(* IEC 61131-3 sources: daoli-st-library/DL_Algo (part 8) *)

(* ---- FB_DL_AutoTuneRelay.st ---- *)
(*
    FB_DL_AutoTuneRelay —— 继电反馈自整定
    ------------------------------------------------------------------
    分类      : DL_Algo / ControlLaw
    前缀      : FB_DL_
    版本      : 1.0.0
    溯源      : 公开学术判据 —— 继电反馈法（Astrom & Hagglund 1984）描述函数
                N(a) = 4d/(pi*a)，含迟滞时 -1/N(a) = -(pi/4d)*sqrt(a^2 - h^2)；
                整定规则取 Ziegler-Nichols 与 Astrom-Hagglund 公开文本；
                只借公开公式与规则常数（属公共知识），测量闸门、状态机、引脚契约与
                码位 100% 自有；clean-room 重写，未复制任何闭源厂商源码
    平台      : 纯 IEC 61131-3，CODESYS V3.5+ / TwinCAT 3 / InoProShop 通用
    作者      : 道莅代码库 · PLC编程专家（R19）
    ------------------------------------------------------------------
    功能说明  : 把 ±d 继电（可带迟滞 h）接入回路，等振幅稳定后测极限振荡周期 Tu 与幅值 a，
                按公开描述函数算临界增益 Ku，再按选定规则给出 Kp / Ti / Td。
                本件不闭环控制，只输出 bRelayOut（接上层手动通道）与整定结果。
                核心防御：① 继电幅值非正/非有限即故障级 2A10（d = 0 时 Ku = 0，结果无意义）；
                ② 迟滞不小于实测幅值时拒绝出结果（描述函数分母为零/虚数，Ku 不可定义）；
                ③ 每半周期采样数不足即故障级 2A11——采样太疏时测出的「振荡」是采样网格
                   产物，不是对象特性（R67 采样密度闸先行）；
                ④ 幅值稳定判据不通过只置信息码继续测，超时才是故障级 2A12；
                ⑤ bAbort 必须撤继电（本件最高危点：不撤则回路一直振荡），且人为中止不置故障。
                说明：继电幅值相对满量程 20% 的工程上限需满量程信息，本件无满量程引脚，
                该上限由调用方在上层保证（头注释留档，不做无法判定的检查）。
    错误码    : 16#0002_2A01 振荡未收敛，继续测量 / 参数超域已钳位——信息级，正常防御
                16#0002_2A02 预留禁用（信息级，不得挪用）
                16#0002_2A10 继电参数非法（d 非正或非有限、h >= a、采样周期越域）——故障级，中止实验并撤继电
                16#0002_2A11 半周期采样密度不足，振荡不可信——故障级，中止实验并撤继电
                16#0002_2A12 超时未收敛 / Ku 不可表示 / 整定规则落 ELSE 兜底——故障级，中止实验并撤继电
    码位总账  : 16#0002_2A01 用 / 16#0002_2A02 预留 ｜ 16#0002_2A10 用 / 16#0002_2A11 用 / 16#0002_2A12 用
    状态机    : E_DL_TuneState（eIdle / eRelay / eMeasure / eDone / eFault）五态，CASE 含 ELSE 兜底，
                ELSE 回 eIdle 并置故障级 2A12；bAbort 沿无条件回 eIdle 且撤继电。
    采样约定  : fbTrigStart / fbTrigAbort / fbTimeout 在本体首部无条件刷新，绝不放入 IF 或 CASE；
                时间基准由 tSampleTime 引脚累加，累加前用比较式预判溢出（不靠回绕兜底）；
                整定规则按公开文本：ZN-P 0.5Ku；ZN-PI 0.45Ku / Tu*1.2^-1；ZN-PID 0.6Ku / Tu/2 / Tu/8；
                AH 无超调 0.2Ku / Tu/2 / Tu/3。
    修订记录  : 2026-11-16 v1.0.0 首次入库（R19）
*)

(*
    枚举 : E_DL_TuneRule —— 整定规则（本文件为全库唯一属主）
*)
TYPE E_DL_TuneRule :
(
    eZnP           := 0,                      // Ziegler-Nichols 纯比例规则 / Ziegler-Nichols proportional rule
    eZnPi          := 1,                      // Ziegler-Nichols 比例积分规则 / Ziegler-Nichols PI rule
    eZnPid         := 2,                      // Ziegler-Nichols 比例积分微分规则 / Ziegler-Nichols PID rule
    eAhNoOvershoot := 3                       // Astrom-Hagglund 无超调规则 / Astrom-Hagglund no overshoot rule
);
END_TYPE

(*
    枚举 : E_DL_TuneState —— 自整定实验状态（本文件为全库唯一属主）
*)
TYPE E_DL_TuneState :
(
    eIdle    := 0,                            // 空闲：继电输出撤销 / idle, relay output withdrawn
    eRelay   := 1,                            // 施加继电，等待首个翻转 / relay applied, waiting for the first flip
    eMeasure := 2,                            // 收集中：测幅值与半周期 / measuring amplitude and half periods
    eDone    := 3,                            // 完成：结果有效 / done, results valid
    eFault   := 4                             // 故障：实验中止 / fault, experiment aborted
);
END_TYPE

FUNCTION_BLOCK FB_DL_AutoTuneRelay
VAR_INPUT
    bEnable           : BOOL;                 // 使能，FALSE 中止实验并撤继电 / enable, FALSE aborts the experiment and withdraws the relay
    bStart            : BOOL;                 // 启动，上升沿启动实验（运行中忽略）/ start, rising edge begins the experiment, ignored while running
    bAbort            : BOOL;                 // 中止，上升沿中止并回 eIdle（不置故障）/ abort, rising edge aborts back to idle without raising a fault
    fPv               : REAL := 0.0;          // 过程测量（被控量）[用户单位] / process measurement [user unit]
    fSp               : REAL := 0.0;          // 目标值，实验围绕此点进行 [用户单位] / setpoint the experiment oscillates around [user unit]
    fRelayAmp         : REAL := 5.0;          // 继电幅值 d [用户单位]，必须 > 0 / relay amplitude d [user unit], must be > 0
    fRelayHyst        : REAL := 0.2;          // 继电迟滞 h [用户单位]，范围 0.0~fRelayAmp（含等号即非法）/ relay hysteresis h [user unit], 0.0~fRelayAmp, equality is illegal
    uCyclesRequired   : UINT := 4;            // 需要观察的完整振荡周期数 [周期]，范围 2~20 / number of full cycles to observe [cycle], range 2~20
    uMinSamplesPerHalf : UINT := 6;           // 每半周期最少采样数 [拍]，范围 4~100 / minimum samples per half period [scan], range 4~100
    tMaxDuration      : TIME := T#300S;       // 实验总超时 [ms]，范围 10 s~2 h / experiment timeout [ms], range 10 s~2 h
    fStabTolPercent   : REAL := 2.0;          // 幅值稳定判据：前后半窗均值差百分比上限 [%]，范围 0.1~20.0 / amplitude stability tolerance [%], range 0.1~20.0
    eRule             : E_DL_TuneRule := eZnPid; // 整定规则 / tuning rule
    tSampleTime       : TIME := T#100MS;      // 采样周期 [ms]，范围 1~10000 / sample time [ms], range 1~10000
END_VAR
VAR_OUTPUT
    bRelayOut         : BOOL;                 // 继电输出（TRUE = 加 +d），接上层手动通道 / relay output, TRUE adds plus d, wired to the manual channel
    bBusy             : BOOL;                 // 实验进行中 / experiment running
    bDone             : BOOL;                 // 完成（单周期脉冲，结果有效）/ done, single-cycle pulse with valid results
    fOscAmp           : REAL;                 // 测得振荡幅值 a [用户单位] / measured oscillation amplitude a [user unit]
    tUltPeriod        : TIME;                 // 测得极限周期 Tu [ms] / measured ultimate period Tu [ms]
    fUltGain          : REAL;                 // 临界增益 Ku [无量纲] / ultimate gain Ku [dimensionless]
    fKp               : REAL;                 // 整定比例增益 [无量纲] / tuned proportional gain [dimensionless]
    fTi               : REAL;                 // 整定积分时间 [s]，0 表示纯 P / tuned integral time [s], zero means pure P
    fTd               : REAL;                 // 整定微分时间 [s]，0 表示无微分 / tuned derivative time [s], zero means no derivative
    uCycleDone        : UINT;                 // 已完成的有效振荡周期数 [周期] / completed valid cycles [cycle]
    eErr              : UDINT;                // 错误码，0=正常 / error id, 0=ok
    bError            : BOOL;                 // 故障标志，eErr 为故障级时 TRUE / error flag, TRUE on fault-level eErr
    bValid            : BOOL;                 // 结果是否可用 / results valid flag
END_VAR
VAR
    eState            : E_DL_TuneState := eIdle; // 状态机当前态 / current state machine state
    fbTrigStart       : R_TRIG;               // 启动沿实例，本体首部无条件刷新 / start edge instance, refreshed unconditionally
    fbTrigAbort       : R_TRIG;               // 中止沿实例，本体首部无条件刷新 / abort edge instance, refreshed unconditionally
    fbTimeout         : TON;                  // 实验总超时实例，本体首部无条件刷新 / total timeout instance, refreshed unconditionally
    bRelayPrev        : BOOL;                 // 上一拍继电输出，翻转检测用 / previous relay output for flip detection
    fPeakHi           : REAL;                 // 本半周期上峰值 [用户单位] / upper peak of the current half period [user unit]
    fPeakLo           : REAL;                 // 本半周期下峰值 [用户单位] / lower peak of the current half period [user unit]
    tNow              : TIME;                 // 实验内累计时间 [ms] / accumulated experiment time [ms]
    tEdgeLast         : TIME;                 // 上一次翻转的时刻 [ms] / time of the previous flip [ms]
    tHalf             : TIME;                 // 最近一个半周期长度 [ms] / most recent half period length [ms]
    tHalfPrev         : TIME;                 // 上一个半周期长度 [ms] / previous half period length [ms]
    uHalfCount        : UINT;                 // 已采集的半周期数 [个] / collected half periods [count]
    fAmpSum1          : REAL;                 // 第一窗幅值累计 [用户单位] / first window amplitude sum [user unit]
    fAmpSum2          : REAL;                 // 第二窗幅值累计 [用户单位] / second window amplitude sum [user unit]
    uAmpCnt1          : UINT;                 // 第一窗样本数 [个] / first window sample count [count]
    uAmpCnt2          : UINT;                 // 第二窗样本数 [个] / second window sample count [count]
    fHalfAmp          : REAL;                 // 单个半周期的幅值 [用户单位] / amplitude of one half period [user unit]
    fMean1            : REAL;                 // 第一窗均值 [用户单位] / first window mean [user unit]
    fMean2            : REAL;                 // 第二窗均值 [用户单位] / second window mean [user unit]
    fRelAmp           : REAL;                 // 幅值相对偏差 [无量纲] / relative amplitude deviation [dimensionless]
    fStabTolEff       : REAL;                 // 钳位后的稳定容差 [%] / clamped stability tolerance [%]
    fCyclesEff        : REAL;                 // 钳位后的周期数（REAL 形态，除法用）/ clamped cycle count in REAL form, used for division
    fHystEff          : REAL;                 // 钳位后的继电迟滞 [用户单位] / clamped relay hysteresis [user unit]
    fKuL              : LREAL;                // 临界增益中间量（LREAL 承载）/ ultimate gain intermediate carried in LREAL
    fAmpL             : LREAL;                // 幅值中间量（LREAL 承载）/ amplitude intermediate carried in LREAL
    fHystL            : LREAL;                // 迟滞中间量（LREAL 承载）/ hysteresis intermediate carried in LREAL
    fDenL             : LREAL;                // 描述函数分母（LREAL 承载）/ describing function denominator in LREAL
    fTuSec            : REAL;                 // 极限周期的秒值 [s] / ultimate period in seconds [s]
    nSampHalf         : DINT;                 // 单半周期采样数 [拍] / samples in one half period [scan]
    nDtMs             : DINT;                 // 采样周期毫秒整数 [ms] / sample time in integer milliseconds [ms]
    uNeedHalf         : UINT;                 // 需要采集的半周期总数 [个] / required half periods [count]
    bNonFin           : BOOL;                 // 输入非有限判定标志 / non-finite input flag
    bCollect          : BOOL;                 // 本拍完成一次有效半周期采集 / a valid half period was collected in this cycle
    uMinSampEff       : UINT;                 // 钳位后的每半周期最少采样数 [拍] / clamped minimum samples per half [scan]
END_VAR
VAR CONSTANT
    DL_AT_MIN_CYCLES    : UINT := 2;          // 周期数下限 [周期] / cycle count lower bound [cycle]
    DL_AT_MAX_CYCLES    : UINT := 20;         // 周期数上限 [周期] / cycle count upper bound [cycle]
    DL_AT_MIN_SAMPLES   : UINT := 4;          // 每半周期采样数下限 [拍] / samples per half lower bound [scan]
    DL_AT_MAX_SAMPLES   : UINT := 100;        // 每半周期采样数上限 [拍] / samples per half upper bound [scan]
    DL_AT_PI            : REAL := 3.14159265; // 圆周率（公开常数）[无量纲] / pi, a public constant [dimensionless]
    DL_AT_FOUR          : LREAL := 4.0;       // 描述函数分子常数 [无量纲] / describing function numerator constant [dimensionless]
    DL_AT_DT_MAX        : TIME := T#10S;      // 采样周期上限 [ms] / sample time upper bound [ms]
    DL_AT_DT_MIN        : TIME := T#1MS;      // 采样周期下限 [ms] / sample time lower bound [ms]
    DL_AT_TIME_MAX      : TIME := T#24H;      // 实验内累计时间饱和值 [ms] / accumulated time saturation [ms]
    DL_AT_TOL_MIN       : REAL := 0.1;        // 稳定容差下限 [%] / stability tolerance lower bound [%]
    DL_AT_TOL_MAX       : REAL := 20.0;       // 稳定容差上限 [%] / stability tolerance upper bound [%]
    DL_FLOAT_EPS        : REAL := 1.0E-6;     // 浮点判等容差 [无量纲] / float equality tolerance [dimensionless]
    DL_AT_PERCENT       : REAL := 100.0;      // 百分比换算因子 [%] / percent conversion factor [%]
    DL_AT_TWO           : REAL := 2.0;        // 二值常量，周期与半周期换算用 [无量纲] / two, used to convert half periods into periods
    DL_AT_ZN_P_K        : REAL := 0.5;        // ZN 纯 P 规则增益系数 [无量纲] / ZN P rule gain factor [dimensionless]
    DL_AT_ZN_PI_K       : REAL := 0.45;       // ZN PI 规则增益系数 [无量纲] / ZN PI rule gain factor [dimensionless]
    DL_AT_ZN_PI_TI      : REAL := 1.2;        // ZN PI 规则积分时间除数 [无量纲] / ZN PI integral time divisor [dimensionless]
    DL_AT_ZN_PID_K      : REAL := 0.6;        // ZN PID 规则增益系数 [无量纲] / ZN PID rule gain factor [dimensionless]
    DL_AT_ZN_PID_TI     : REAL := 2.0;        // ZN PID 规则积分时间除数 [无量纲] / ZN PID integral time divisor [dimensionless]
    DL_AT_ZN_PID_TD     : REAL := 8.0;        // ZN PID 规则微分时间除数 [无量纲] / ZN PID derivative time divisor [dimensionless]
    DL_AT_AH_K          : REAL := 0.2;        // AH 无超调规则增益系数 [无量纲] / AH no overshoot gain factor [dimensionless]
    DL_AT_AH_TI         : REAL := 2.0;        // AH 无超调规则积分时间除数 [无量纲] / AH integral time divisor [dimensionless]
    DL_AT_AH_TD         : REAL := 3.0;        // AH 无超调规则微分时间除数 [无量纲] / AH derivative time divisor [dimensionless]
    DL_AT_MS_PER_S      : REAL := 1000.0;     // 毫秒到秒换算因子 [ms/s] / milliseconds per second [ms/s]
    DL_AT_ZERO          : REAL := 0.0;        // 零值常量，避免裸字面量 [无量纲] / zero constant, avoids a bare literal [dimensionless]
    DL_AT_ZERO_L        : LREAL := 0.0;       // LREAL 零值常量 [无量纲] / LREAL zero constant [dimensionless]
    DL_AT_KU_MAX        : LREAL := 1.0E30;    // 临界增益可表示上限 [无量纲] / representable upper bound of the critical gain [dimensionless]
    DL_AT_INF_GUARD     : REAL := 1.0E38;     // 非有限幅值判定阈值 [无量纲] / non-finite magnitude guard [dimensionless]
    DL_AT_TWO_I         : INT := 2;           // 整形二值常量，半周期转周期用 [无量纲] / integer two, converts half periods into periods
    DL_AT_TWO_U         : UINT := 2;          // 无符号二值常量，半周期数折周期数用 [无量纲] / unsigned two, folds half periods into cycles
END_VAR

// 段 1｜边沿与定时器实例无条件周期刷新（红线：严禁放入条件分支）/ segment 1, unconditional refresh
fbTrigStart(CLK := bStart);
fbTrigAbort(CLK := bAbort);
fbTimeout(IN := (eState = eRelay) OR (eState = eMeasure), PT := tMaxDuration); // 只有实验期计时 / the timer runs only during the experiment

// 段 2｜输出与错误状态预置（结果量保持，bDone 为单周期脉冲）/ segment 2, preset outputs and status
bDone := FALSE;                               // 脉冲先清 / clear the pulse first
eErr := 0;                                    // 预置无错误 / preset no error
bError := FALSE;                              // 预置无故障 / preset no fault
bValid := FALSE;                              // 预置结果不可用 / preset results invalid
bCollect := FALSE;                            // 预置本拍无采集 / preset no collection in this cycle
bBusy := (eState = eRelay) OR (eState = eMeasure); // 忙标志由状态导出 / the busy flag derives from the state

// 段 3｜输入非有限闸：直接落故障态并撤继电 / segment 3, non-finite gate
bNonFin := (fPv <> fPv) OR (fSp <> fSp) OR (fRelayAmp <> fRelayAmp) OR (fRelayHyst <> fRelayHyst); // 非有限判定 / non-finite detection
IF bNonFin THEN
    eErr := 16#0002_2A10;                     // 继电参数非法故障码 / illegal relay parameter fault id
    bError := TRUE;                           // 置故障标志 / raise the error flag
    eState := eFault;                         // 落故障态 / enter the fault state
    bRelayOut := FALSE;                       // 撤继电，绝不留在振荡状态 / withdraw the relay, never leave the loop oscillating
    RETURN;                                   // 故障级提前返回 / early return on fault
END_IF

// 段 4｜中止沿：人为中止不置故障，但必须撤继电 / segment 4, abort edge withdraws the relay without a fault
IF fbTrigAbort.Q THEN
    eState := eIdle;                          // 回空闲态 / back to idle
    bRelayOut := FALSE;                       // 撤继电（本件最高危点）/ withdraw the relay, the most critical point of this block
    bBusy := FALSE;                           // 忙标志撤销 / drop the busy flag
    RETURN;                                   // 中止即出口 / abort is the exit
END_IF

// 段 5｜失能闸：失能同样撤继电 / segment 5, enable gate
IF NOT bEnable THEN
    eState := eIdle;                          // 回空闲态 / back to idle
    bRelayOut := FALSE;                       // 撤继电 / withdraw the relay
    bBusy := FALSE;                           // 忙标志撤销 / drop the busy flag
    RETURN;                                   // 失能即出口 / disabled is the exit
END_IF

// 段 6｜参数域钳位（周期数、采样数、容差、迟滞、超时）/ segment 6, parameter domain clamp
IF (uCyclesRequired < DL_AT_MIN_CYCLES) THEN
    uNeedHalf := DL_AT_MIN_CYCLES;            // 周期数下限钳位 / clamp at the lower cycle count
    eErr := 16#0002_2A01;                     // 信息级：参数超域已钳位 / info level, the parameter was clamped
ELSIF (uCyclesRequired > DL_AT_MAX_CYCLES) THEN
    uNeedHalf := DL_AT_MAX_CYCLES;            // 周期数上限钳位 / clamp at the upper cycle count
    eErr := 16#0002_2A01;                     // 信息级：参数超域已钳位 / info level, the parameter was clamped
ELSE
    uNeedHalf := uCyclesRequired;             // 域内直接用 / in-domain value
END_IF
fCyclesEff := UINT_TO_REAL(uNeedHalf);        // 周期数 REAL 形态，除法前保证非零 / REAL form of the cycle count, nonzero by construction
fStabTolEff := MIN(MAX(fStabTolPercent, DL_AT_TOL_MIN), DL_AT_TOL_MAX); // 稳定容差收敛到 0.1~20.0 % / converge the tolerance into 0.1~20.0 %
fHystEff := MIN(MAX(fRelayHyst, DL_AT_ZERO), fRelayAmp); // 迟滞收敛到 0.0~d / converge the hysteresis into 0.0~d
IF uMinSamplesPerHalf < DL_AT_MIN_SAMPLES THEN
    uMinSampEff := DL_AT_MIN_SAMPLES;         // 采样数下限钳位 / clamp at the lower sample count
    eErr := 16#0002_2A01;                     // 信息级：参数超域已钳位 / info level, the parameter was clamped
ELSIF uMinSamplesPerHalf > DL_AT_MAX_SAMPLES THEN
    uMinSampEff := DL_AT_MAX_SAMPLES;         // 采样数上限钳位 / clamp at the upper sample count
    eErr := 16#0002_2A01;                     // 信息级：参数超域已钳位 / info level, the parameter was clamped
ELSE
    uMinSampEff := uMinSamplesPerHalf;        // 域内直接用 / in-domain value
END_IF
nDtMs := TIME_TO_DINT(tSampleTime);           // 采样周期整数毫秒 [ms] / sample time in integer milliseconds [ms]

// 段 7｜启动前提闸（幅值、采样周期、超时、采样数）/ segment 7, start preconditions
IF fbTrigStart.Q AND ((eState = eIdle) OR (eState = eDone) OR (eState = eFault)) THEN
    IF (fRelayAmp <= DL_FLOAT_EPS) OR (ABS(fRelayAmp) > DL_AT_INF_GUARD)
       OR (tSampleTime < DL_AT_DT_MIN) OR (tSampleTime > DL_AT_DT_MAX) THEN
        eErr := 16#0002_2A10;                 // 继电幅值为 0 时 Ku 恒 0，整定结果无意义 / a zero amplitude makes Ku zero and the result meaningless
        bError := TRUE;                       // 置故障标志 / raise the error flag
        eState := eFault;                     // 落故障态 / enter the fault state
        bRelayOut := FALSE;                   // 撤继电 / withdraw the relay
        RETURN;                               // 故障级提前返回 / early return on fault
    END_IF
    // 段 8｜实验现场复位并进入继电器相 / segment 8, reset the experiment context and start the relay phase
    eState := eRelay;                         // 进入继电器相 / enter the relay phase
    tNow := T#0S;                             // 累计时间清零 / clear the accumulated time
    tEdgeLast := T#0S;                        // 翻转时刻清零 / clear the flip timestamp
    tHalf := T#0S;                            // 半周期清零 / clear the half period
    tHalfPrev := T#0S;                        // 上一半周期清零 / clear the previous half period
    uHalfCount := 0;                          // 半周期计数清零 / clear the half period counter
    fAmpSum1 := DL_AT_ZERO;                   // 第一窗清零 / clear the first window
    fAmpSum2 := DL_AT_ZERO;                   // 第二窗清零 / clear the second window
    uAmpCnt1 := 0;                            // 第一窗计数清零 / clear the first window count
    uAmpCnt2 := 0;                            // 第二窗计数清零 / clear the second window count
    fPeakHi := fPv;                           // 峰值基准取当前测量 / seed the peaks from the current measurement
    fPeakLo := fPv;                           // 峰值基准取当前测量 / seed the peaks from the current measurement
    bRelayPrev := FALSE;                      // 翻转检测基准复位 / reset the flip reference
    bRelayOut := (fPv < fSp);                 // 初始继电方向：低于目标则加 +d / initial relay direction, add plus d below the setpoint
END_IF

// 段 9｜时间累加（比较式预判溢出，不靠回绕兜底）/ segment 9, accumulated time with a comparison overflow guard
IF ((eState = eRelay) OR (eState = eMeasure)) AND (tNow < (DL_AT_TIME_MAX - tSampleTime)) THEN
    tNow := tNow + tSampleTime;               // 累计实验时间 [ms] / accumulate the experiment time [ms]
END_IF

// 段 10｜状态机（含 ELSE 兜底）/ segment 10, state machine with ELSE fallback
CASE eState OF
    eIdle:
        bRelayOut := FALSE;                   // 空闲态无继电输出 / no relay output while idle
        bBusy := FALSE;                       // 空闲态不忙 / not busy while idle

    eRelay:
        // 段 11｜继电翻转（带迟滞）：低于 Sp−h 加 +d，高于 Sp+h 加 −d，带内保持 / segment 11, relay switching with hysteresis
        IF fPv < (fSp - fHystEff) THEN
            bRelayOut := TRUE;                // 低于下界，加正幅值 / below the lower band, apply plus d
        ELSIF fPv > (fSp + fHystEff) THEN
            bRelayOut := FALSE;               // 高于上界，加负幅值 / above the upper band, apply minus d
        END_IF
        fPeakHi := MAX(fPeakHi, fPv);         // 跟踪上峰值 / track the upper peak
        fPeakLo := MIN(fPeakLo, fPv);         // 跟踪下峰值 / track the lower peak
        IF bRelayOut <> bRelayPrev THEN
            bRelayPrev := bRelayOut;          // 记录新方向 / remember the new direction
            tEdgeLast := tNow;                // 记录首个翻转时刻 / remember the first flip instant
            fPeakHi := fPv;                   // 峰值重新播种 / reseed the peaks
            fPeakLo := fPv;                   // 峰值重新播种 / reseed the peaks
            eState := eMeasure;               // 首个翻转即进入测量相 / the first flip enters the measuring phase
        END_IF

    eMeasure:
        // 段 12｜同段内继续翻转判定 / segment 12, continued switching inside the measuring phase
        IF fPv < (fSp - fHystEff) THEN
            bRelayOut := TRUE;                // 低于下界，加正幅值 / below the lower band, apply plus d
        ELSIF fPv > (fSp + fHystEff) THEN
            bRelayOut := FALSE;               // 高于上界，加负幅值 / above the upper band, apply minus d
        END_IF
        fPeakHi := MAX(fPeakHi, fPv);         // 跟踪上峰值 / track the upper peak
        fPeakLo := MIN(fPeakLo, fPv);         // 跟踪下峰值 / track the lower peak

        // 段 13｜翻转沿：结算一个半周期的幅值与长度，并做采样密度闸 / segment 13, settle one half period and check the sample density
        IF bRelayOut <> bRelayPrev THEN
            tHalfPrev := tHalf;               // 保留上一个半周期 / keep the previous half period
            tHalf := tNow - tEdgeLast;        // 本半周期长度 [ms] / this half period length [ms]
            tEdgeLast := tNow;                // 更新翻转时刻 / update the flip instant
            fHalfAmp := (fPeakHi - fPeakLo) / DL_AT_TWO; // 半周期幅值 [用户单位] / half period amplitude [user unit]
            fPeakHi := fPv;                   // 峰值重新播种 / reseed the peaks
            fPeakLo := fPv;                   // 峰值重新播种 / reseed the peaks
            bRelayPrev := bRelayOut;          // 记录新方向 / remember the new direction
            IF nDtMs > 0 THEN
                nSampHalf := TIME_TO_DINT(tHalf) / nDtMs; // 半周期采样数（整数除法，除子已判非零）/ samples per half, integer division with a guarded divisor
                IF nSampHalf < UINT_TO_DINT(uMinSampEff) THEN
                    eErr := 16#0002_2A11;     // 采样过疏，测到的振荡是采样网格产物 / too sparse, the measured oscillation is a sampling artefact
                    bError := TRUE;           // 置故障标志 / raise the error flag
                    eState := eFault;         // 落故障态 / enter the fault state
                    bRelayOut := FALSE;       // 撤继电 / withdraw the relay
                    RETURN;                   // 故障级提前返回 / early return on fault
                END_IF
            END_IF
            uHalfCount := uHalfCount + 1;     // 半周期计数加一 / increment the half period counter
            bCollect := TRUE;                 // 标记本拍完成采集 / flag the collection in this cycle
            IF uAmpCnt1 < uNeedHalf THEN
                fAmpSum1 := fAmpSum1 + fHalfAmp; // 第一窗累计幅值 / accumulate into the first window
                uAmpCnt1 := uAmpCnt1 + 1;     // 第一窗计数加一 / increment the first window count
            ELSE
                fAmpSum2 := fAmpSum2 + fHalfAmp; // 第二窗累计幅值 / accumulate into the second window
                uAmpCnt2 := uAmpCnt2 + 1;     // 第二窗计数加一 / increment the second window count
            END_IF
            uCycleDone := uHalfCount / DL_AT_TWO_U; // 已完成的有效周期数由半周期数折半 / completed cycles folded from the half period count
        END_IF

        // 段 14｜两窗齐备后判稳定：不稳只置信息码继续测，超时才是故障 / segment 14, stability check
        IF bCollect AND (uAmpCnt1 >= uNeedHalf) AND (uAmpCnt2 >= uNeedHalf) THEN
            fMean1 := fAmpSum1 / fCyclesEff;  // 第一窗均值，除子为周期数（≥ 2）/ first window mean, the divisor is at least two
            fMean2 := fAmpSum2 / fCyclesEff;  // 第二窗均值 / second window mean
            IF ((fMean1 + fMean2) * DL_AT_TWO) > DL_FLOAT_EPS THEN
                fRelAmp := ABS(fMean1 - fMean2) / ((fMean1 + fMean2) / DL_AT_TWO) * DL_AT_PERCENT; // 相对偏差 [%] / relative deviation [%]
            ELSE
                fRelAmp := DL_AT_PERCENT;     // 幅值近零时视为完全不一致 / a near zero amplitude counts as fully inconsistent
            END_IF
            IF fRelAmp > fStabTolEff THEN
                eErr := 16#0002_2A01;         // 信息级：振荡未收敛，清窗继续测 / info level, not converged, clear the windows and continue
                fAmpSum1 := DL_AT_ZERO;       // 清第一窗（重新收集）/ clear the first window and collect again
                fAmpSum2 := DL_AT_ZERO;       // 清第二窗 / clear the second window
                uAmpCnt1 := 0;                // 清第一窗计数 / clear the first window count
                uAmpCnt2 := 0;                // 清第二窗计数 / clear the second window count
            ELSE
                // 段 15｜临界增益：Ku = 4d / (pi·sqrt(a^2 − h^2))，含迟滞时退化为 4d/(pi·a) / segment 15, critical gain
                fOscAmp := (fMean1 + fMean2) / DL_AT_TWO; // 振荡幅值取两窗均值 [用户单位] / amplitude as the mean of both windows [user unit]
                tUltPeriod := tHalfPrev * DL_AT_TWO_I;  // 极限周期取最近半周期×2 [ms] / ultimate period as twice the latest half period [ms]
                fTuSec := DINT_TO_REAL(TIME_TO_DINT(tUltPeriod)) / DL_AT_MS_PER_S; // 极限周期秒值 [s] / ultimate period in seconds [s]
                IF fHystEff >= fOscAmp THEN
                    eErr := 16#0002_2A10;     // 迟滞不小于实测幅值，描述函数分母为零/虚数 / hysteresis not narrower than the amplitude makes the denominator zero or imaginary
                    bError := TRUE;           // 置故障标志 / raise the error flag
                    eState := eFault;         // 落故障态 / enter the fault state
                    bRelayOut := FALSE;       // 撤继电 / withdraw the relay
                    RETURN;                   // 故障级提前返回 / early return on fault
                END_IF
                fAmpL := REAL_TO_LREAL(fOscAmp);   // 幅值升位到 LREAL / widen the amplitude to LREAL
                fHystL := REAL_TO_LREAL(fHystEff); // 迟滞升位到 LREAL / widen the hysteresis to LREAL
                fDenL := fAmpL * fAmpL - fHystL * fHystL; // a^2 − h^2（含迟滞描述函数分母）/ squared amplitude minus squared hysteresis
                IF fDenL <= DL_AT_ZERO_L THEN
                    eErr := 16#0002_2A12;     // 分母非正，Ku 不可表示 / the denominator is not positive, Ku is not representable
                    bError := TRUE;           // 置故障标志 / raise the error flag
                    eState := eFault;         // 落故障态 / enter the fault state
                    bRelayOut := FALSE;       // 撤继电 / withdraw the relay
                    RETURN;                   // 故障级提前返回 / early return on fault
                END_IF
                fKuL := DL_AT_FOUR * REAL_TO_LREAL(fRelayAmp) / (REAL_TO_LREAL(DL_AT_PI) * SQRT(fDenL)); // 临界增益（LREAL 中间量）/ critical gain carried in LREAL
                IF (fKuL <> fKuL) OR (fKuL <= DL_AT_ZERO_L) OR (fKuL > DL_AT_KU_MAX) THEN
                    eErr := 16#0002_2A12;     // Ku 不可表示 / Ku is not representable
                    bError := TRUE;           // 置故障标志 / raise the error flag
                    eState := eFault;         // 落故障态 / enter the fault state
                    bRelayOut := FALSE;       // 撤继电 / withdraw the relay
                    RETURN;                   // 故障级提前返回 / early return on fault
                END_IF
                fUltGain := LREAL_TO_REAL(fKuL);   // 回落到 REAL 输出 / narrow back to REAL for the output
                // 段 16｜整定规则（公开文本常数，CASE 含 ELSE 兜底）/ segment 16, tuning rules with ELSE fallback
                CASE eRule OF
                    eZnP:
                        fKp := DL_AT_ZN_P_K * fUltGain;              // 纯比例：Kp = 0.5·Ku / proportional only
                        fTi := DL_AT_ZERO;                           // 纯 P 无积分 / pure P has no integral
                        fTd := DL_AT_ZERO;                           // 纯 P 无微分 / pure P has no derivative
                    eZnPi:
                        fKp := DL_AT_ZN_PI_K * fUltGain;             // PI：Kp = 0.45·Ku / PI gain
                        fTi := fTuSec / DL_AT_ZN_PI_TI;              // PI：Ti = Tu / 1.2 [s] / PI integral time
                        fTd := DL_AT_ZERO;                           // PI 无微分 / PI has no derivative
                    eZnPid:
                        fKp := DL_AT_ZN_PID_K * fUltGain;            // PID：Kp = 0.6·Ku / PID gain
                        fTi := fTuSec / DL_AT_ZN_PID_TI;             // PID：Ti = Tu / 2 [s] / PID integral time
                        fTd := fTuSec / DL_AT_ZN_PID_TD;             // PID：Td = Tu / 8 [s] / PID derivative time
                    eAhNoOvershoot:
                        fKp := DL_AT_AH_K * fUltGain;                // 无超调：Kp = 0.2·Ku / no overshoot gain
                        fTi := fTuSec / DL_AT_AH_TI;                 // 无超调：Ti = Tu / 2 [s] / no overshoot integral time
                        fTd := fTuSec / DL_AT_AH_TD;                 // 无超调：Td = Tu / 3 [s] / no overshoot derivative time
                ELSE
                    eErr := 16#0002_2A12;                            // 故障级：非法规则兜底 / fault level, illegal rule fallback
                    bError := TRUE;                                  // 置故障标志 / raise the error flag
                    eState := eFault;                                // 落故障态 / enter the fault state
                    bRelayOut := FALSE;                              // 撤继电 / withdraw the relay
                    RETURN;                                          // 故障级提前返回 / early return on fault
                END_CASE
                eState := eDone;              // 结果产出，进入完成态 / results produced, enter the done state
                bDone := TRUE;                // 单周期完成脉冲 / single-cycle done pulse
                bRelayOut := FALSE;           // 完成后必须撤继电 / withdraw the relay once finished
                bValid := TRUE;               // 结果可用 / results are valid
                bBusy := FALSE;               // 实验结束 / the experiment is finished
            END_IF
        END_IF

    eDone:
        bRelayOut := FALSE;                   // 完成态保持无继电输出 / no relay output in the done state
        bValid := TRUE;                       // 结果保持可用 / results stay valid
        bBusy := FALSE;                       // 不忙 / not busy

    eFault:
        bRelayOut := FALSE;                   // 故障态撤继电 / withdraw the relay in the fault state
        bBusy := FALSE;                       // 不忙 / not busy

ELSE
    eErr := 16#0002_2A12;                     // 故障级：非法状态兜底 / fault level, illegal state fallback
    bError := TRUE;                           // 置故障标志 / raise the error flag
    eState := eIdle;                          // 回空闲态 / fall back to idle
    bRelayOut := FALSE;                       // 撤继电，绝不留振荡 / withdraw the relay, never leave the loop oscillating
END_CASE

// 段 17｜超时闸：只有实验期有效，超时即故障并撤继电 / segment 17, timeout gate
IF fbTimeout.Q AND ((eState = eRelay) OR (eState = eMeasure)) THEN
    eErr := 16#0002_2A12;                     // 超时未收敛故障码 / timeout without convergence fault id
    bError := TRUE;                           // 置故障标志 / raise the error flag
    eState := eFault;                         // 落故障态 / enter the fault state
    bRelayOut := FALSE;                       // 撤继电 / withdraw the relay
END_IF
END_FUNCTION_BLOCK

(* ---- FB_DL_BearingVibTrend.st ---- *)
(*
  Name        : FB_DL_BearingVibTrend
  Category    : DL_Algo
  Version     : 1.0.0
  Purpose     : 轴承振动 RMS 滑窗趋势分级预警：采样触发下把振动 RMS 入环形窗，按窗内均值与峰值对 ISO 10816 三档门槛（良好/注意/报警）分级；/ Bearing vibration RMS sliding-window trend: RMS samples enter a ring window, graded against ISO 10816 three-band thresholds by window mean and peak
  溯源        : 借 t2-1-lgf-measurement 的分类/参数域组织，clean-room 实现
  Boundary    : ① 组态闸：窗长域 4..32 / 注意与报警门槛须正且注意 < 报警 → 锁存故障；
                ② 环窗时间序范式（R194/R205）：_nHead 声明即赋初值 1；窗深变更后回钳 _nHead/_nFill，防越界写与环序破坏；
                ③ 非有限 RMS 该次不入样（拒收计数 bSampleRej 供诊断），不污染统计；
                ④ 分级判据全部 >= 阈值直比（阈值来自组态，非浮点等值比较）；
                ⑤ 本件为趋势诊断层，不停机不联锁（属主边界）。
*)
TYPE E_DL_BvtState :
(
    eIdle  := 0,                             (* 未使能 / Disabled *)
    eMon   := 10,                            (* 趋势监视运行 / Monitoring *)
    eFault := 90                             (* 故障锁存相 / Fault latched *)
);
END_TYPE

TYPE E_DL_BvtCause :
(
    eNone       := 0,                        (* 无故障成因 / No cause *)
    eCfgIllegal := 1,                        (* 组态非法：窗长/门槛越域 / Illegal config *)
    ePhaseBad   := 2                         (* 非法相位兜底 / Illegal phase fallback *)
);
END_TYPE

FUNCTION_BLOCK FB_DL_BearingVibTrend
VAR_INPUT
    fVibRms   : REAL := 0.0;                 (* 振动速度 RMS 实测 [mm/s] / Vibration velocity RMS *)
    bSample   : BOOL := FALSE;               (* 采样触发脉冲（上升沿采一个样本）[-] / Sample trigger pulse *)
    nWinLen   : INT := 16;                   (* 滑窗深度，域 4..32 [点] / Window depth, 4..32 *)
    fThGood   : REAL := 2.8;                 (* ISO 10816 良好档上限（A/B 分界），域 > 0 [mm/s] / Good-band limit *)
    fThAlert  : REAL := 7.1;                 (* ISO 10816 报警档下限（C/D 分界），域 > 注意档 [mm/s] / Alarm-band limit *)
    bEnable   : BOOL := TRUE;                (* 监视使能 [-] / Enable *)
    bReset    : BOOL := FALSE;               (* 复位命令，上升沿清窗与预警 [-] / Reset command *)
END_VAR
VAR_OUTPUT
    fRmsMean  : REAL;                        (* 窗内 RMS 均值 [mm/s] / Window mean *)
    fRmsPeak  : REAL;                        (* 窗内 RMS 峰值 [mm/s] / Window peak *)
    nFill     : INT;                         (* 窗内有效样本数 [点] / Valid samples in window *)
    bGood     : BOOL;                        (* 分级：良好档（均值 <= 良好门槛）[-] / Good band *)
    bAlert    : BOOL;                        (* 分级：注意档（未达报警但超良好门槛）[-] / Alert band *)
    bAlarm    : BOOL;                        (* 分级：报警档（峰值或均值 >= 报警门槛）[-] / Alarm band *)
    bSampleRej: BOOL;                        (* 本拍有非有限样本被拒收 [-] / Sample rejected this scan *)
    eState    : E_DL_BvtState;               (* 状态出口 / State outlet *)
    eCause    : E_DL_BvtCause;               (* 故障成因出口（R190 归因唯一） / Fault cause outlet *)
    bError    : BOOL;                        (* 故障锁存标志 [-] / Fault latch flag *)
END_VAR
VAR
    _eState  : E_DL_BvtState := E_DL_BvtState.eIdle;     (* 内部相位（CASE 唯一写入目标） / Internal phase *)
    _eCause  : E_DL_BvtCause := E_DL_BvtCause.eNone;     (* 故障成因锁存量 / Latched cause *)
    rtSample : R_TRIG;                       (* 采样触发沿实例，段 0 无条件调用 / Sample edge instance *)
    rtReset  : R_TRIG;                       (* 复位沿实例，段 0 无条件调用 / Reset edge instance *)
    _bFault  : BOOL;                         (* 故障锁存位 / Latched fault bit *)
    _bCfgBad : BOOL;                         (* 组态非法当拍量 / Illegal config this scan *)
    _bFin    : BOOL;                         (* RMS 有限性当拍量 / RMS finiteness *)
    _aRms    : ARRAY[1..32] OF REAL;         (* 振动 RMS 环形样本数组 [mm/s] / Ring buffer of RMS samples *)
    _nHead   : INT := 1;                     (* 环形写头（声明即赋初值 1，R194 教训） / Ring write head, init 1 *)
    _nFill   : INT;                          (* 环窗已填样本数 [点] / Ring fill count *)
    _nEff    : INT;                          (* 钳位后生效窗深 [点] / Effective window depth *)
    _nIdx    : INT;                          (* 统计游标（每趟重置，R227）[-] / Stats cursor *)
    _fSum    : REAL;                         (* Σx 中间量 [mm/s] / Sum intermediate *)
    _fMeanI  : REAL;                         (* 均值中间量 [mm/s] / Mean intermediate *)
    _fPeakI  : REAL;                         (* 峰值中间量 [mm/s] / Peak intermediate *)
END_VAR
VAR CONSTANT
    DL_BVT_EPS    : REAL := 1.0E-6;          (* 判零容差 [-] / Epsilon *)
    DL_BVT_NMAX   : INT  := 32;              (* 窗容量上限 [点] / Window capacity *)
    DL_BVT_NMIN   : INT  := 4;               (* 窗深下限（保证趋势统计有效）[点] / Window depth lower bound *)
END_VAR

(* —— 段 0：当拍判据派生 + 实例无条件刷新（R228A；R_TRIG 全在段 0，无 IF 包裹） —— *)
_bCfgBad := (nWinLen < DL_BVT_NMIN) OR (nWinLen > DL_BVT_NMAX)                 (* 窗长域闸 / Window-depth gate *)
            OR (fThGood <= DL_BVT_EPS)                                         (* 良好门槛正域闸 / Good-limit gate *)
            OR (fThAlert <= fThGood);                                          (* 报警门槛须大于注意/良好门槛（防档位倒置） / Alarm limit above good limit *)
rtSample(CLK := bSample);                                                      (* 采样沿每拍必调 / Sample edge every scan *)
rtReset(CLK := bReset);                                                        (* 复位沿每拍必调 / Reset edge every scan *)
_bFin := (fVibRms = fVibRms) AND ((fVibRms - fVibRms) = (fVibRms - fVibRms));  (* RMS NaN 自反 + Inf 差判闸 / RMS NaN and Inf gate *)
_nEff := nWinLen;                                                              (* 生效窗深初值 / Effective depth init *)
IF _nEff < DL_BVT_NMIN THEN
    _nEff := DL_BVT_NMIN;                                                      (* 窗深下限钳位 / Lower clamp *)
END_IF
IF _nEff > DL_BVT_NMAX THEN
    _nEff := DL_BVT_NMAX;                                                      (* 窗深上限钳位（R308） / Upper clamp *)
END_IF
IF _nHead > _nEff THEN
    _nHead := 1;                                                               (* 窗深变小后回钳写头（环序重同步，R194/R205） / Re-clamp head after depth shrink *)
END_IF
IF _nFill > _nEff THEN
    _nFill := _nEff;                                                           (* 窗深变小后回钳填充数（防封顶失效） / Re-clamp fill after depth shrink *)
END_IF

(* —— 段 1：单拍量预清零（R107） —— *)
bSampleRej := FALSE;                                                           (* 拒收指示预清 / Reject-sample preset *)
bGood := FALSE;                                                                (* 良好档预清 / Good preset *)
bAlert := FALSE;                                                               (* 注意档预清 / Alert preset *)
bAlarm := FALSE;                                                               (* 报警档预清 / Alarm preset *)

(* —— 段 2：复位沿处理（作用域：清故障 + 清环窗（仅头/填充数与游标，数据域随填充数失效）+ 清出口 + 迁 eIdle，R283 逐项声明） —— *)
IF rtReset.Q THEN
    _bFault := FALSE;                                                          (* 清故障锁存 / Clear fault *)
    _eCause := E_DL_BvtCause.eNone;                                            (* 清成因 / Clear cause *)
    _nHead := 1;                                                               (* 写头回 1（声明同值） / Head back to 1 *)
    _nFill := 0;                                                               (* 清填充数（旧数据随计数失效） / Clear fill *)
    nFill := 0;                                                                (* 清填充数出口 / Clear fill outlet *)
    fRmsMean := 0.0;                                                           (* 清均值出口 / Clear mean outlet *)
    fRmsPeak := 0.0;                                                           (* 清峰值出口 / Clear peak outlet *)
    _eState := E_DL_BvtState.eIdle;                                            (* 迁未使能相 / Back to idle *)
END_IF

(* —— 段 3：组态故障锁存（锁存至复位沿，R189） —— *)
IF _bCfgBad AND NOT _bFault THEN
    _bFault := TRUE;                                                           (* 锁存故障位 / Latch fault *)
    _eCause := E_DL_BvtCause.eCfgIllegal;                                      (* 成因：组态非法 / Cause: illegal config *)
    _eState := E_DL_BvtState.eFault;                                           (* 同步迁故障相 / Migrate to fault *)
END_IF

(* —— 段 4：CASE 主状态机（ELSE 兜底迁 eFault，红线 6） —— *)
CASE _eState OF
    E_DL_BvtState.eIdle:                                                       (* 未使能：不采样 / Disabled *)
        _nFill := 0;                                                           (* 失能清填充数（防隐性回夹） / Clear fill *)
        nFill := 0;                                                            (* 失能清填充数出口 / Clear fill outlet *)
        fRmsMean := 0.0;                                                       (* 失能清均值出口（eIdle/eFault 出口确定值） / Clear mean outlet *)
        fRmsPeak := 0.0;                                                       (* 失能清峰值出口 / Clear peak outlet *)
        IF bEnable AND NOT _bFault THEN
            _eState := E_DL_BvtState.eMon;                                     (* 使能进入监视 / Enter monitoring *)
        END_IF
    E_DL_BvtState.eMon:                                                        (* 监视相：采样入窗 + 统计分级 / Monitoring *)
        IF NOT bEnable THEN
            _eState := E_DL_BvtState.eIdle;                                    (* 失能回未使能 / Back to idle *)
        ELSIF rtSample.Q THEN                                                  (* 采样触发：一次入样 / Sample trigger *)
            IF _bFin THEN                                                      (* 有限样本入窗 / Finite sample accepted *)
                _aRms[_nHead] := fVibRms;                                      (* 环窗写入（下标已由段 0 回钳保证 1.._nEff） / Ring write, index clamped *)
                _nHead := _nHead + 1;                                          (* 写头递进 / Head advance *)
                IF _nHead > _nEff THEN
                    _nHead := 1;                                               (* 写头回卷到 1 / Head wrap to 1 *)
                END_IF
                IF _nFill < _nEff THEN
                    _nFill := _nFill + 1;                                      (* 未满窗则填充数递增 / Fill up to depth *)
                END_IF
                nFill := _nFill;                                               (* 填充数出口镜像 / Fill outlet mirror *)
            ELSE
                bSampleRej := TRUE;                                            (* 非有限样本拒收（边界③） / Reject non-finite *)
            END_IF
            _fSum := 0.0;                                                      (* Σx 预清 / Sum preset *)
            _fPeakI := 0.0;                                                    (* 峰值预清（RMS 恒 >= 0，0 起步安全） / Peak preset *)
            _nIdx := 1;                                                        (* 游标起头（R227） / Cursor reset *)
            WHILE _nIdx <= _nFill DO                                           (* 一趟求 Σx/峰值（下标域 1.._nFill 有界） / One pass for sum and peak *)
                _fSum := _fSum + _aRms[_nIdx];                                 (* Σx [mm/s] / Sum *)
                IF _aRms[_nIdx] > _fPeakI THEN
                    _fPeakI := _aRms[_nIdx];                                   (* 更新峰值 / Update peak *)
                END_IF
                _nIdx := _nIdx + 1;                                            (* 游标递进 / Cursor advance *)
            END_WHILE
            IF _nFill >= DL_BVT_NMIN THEN                                      (* 窗内样本足额才刷新统计与分级 / Grade only with enough samples *)
                _fMeanI := _fSum / DINT_TO_REAL(_nFill);                       (* 均值：除子 _nFill >= 4 无除零 [mm/s] / Mean, divisor >= 4 *)
                fRmsMean := _fMeanI;                                           (* 均值出口 / Mean outlet *)
                fRmsPeak := _fPeakI;                                           (* 峰值出口 / Peak outlet *)
                IF (_fPeakI >= fThAlert) OR (_fMeanI >= fThAlert) THEN
                    bAlarm := TRUE;                                            (* 报警档：峰值或均值达报警门槛 / Alarm band *)
                ELSIF (_fPeakI >= fThGood) OR (_fMeanI >= fThGood) THEN
                    bAlert := TRUE;                                            (* 注意档：超良好门槛未达报警 / Alert band *)
                ELSE
                    bGood := TRUE;                                             (* 良好档：均值与峰值均低于良好门槛 / Good band *)
                END_IF
            END_IF
        END_IF
    E_DL_BvtState.eFault:                                                      (* 故障相：冻结保持末值，仅复位沿出 / Fault *)
        ;                                                                      (* 锁存回放（R28） / Replay from latch *)
    ELSE                                                                       (* 非法相位兜底迁安全态 / Illegal phase fallback *)
        _eState := E_DL_BvtState.eFault;                                       (* 迁故障相 / To fault *)
        _bFault := TRUE;                                                       (* 同步锁存 / Latch *)
        _eCause := E_DL_BvtCause.ePhaseBad;                                    (* 成因：非法相位 / Cause: illegal phase *)
END_CASE

(* —— 段 5：出口映射（bError/eState 同源，R191） —— *)
bError := _bFault;                                                             (* 故障标志镜像 / Fault flag mirror *)
eState := _eState;                                                             (* 状态出口 / State outlet *)
eCause := _eCause;                                                             (* 成因出口 / Cause outlet *)
END_FUNCTION_BLOCK

(* ---- FB_DL_BiasAdaptiveTrim.st ---- *)
(*==============================================================================
 * 组件名称 (Component)  : FB_DL_BiasAdaptiveTrim
 * 所属子库 (Sublibrary) : DL_Algo
 * 当前版本 (Version)    : 1.0.0
 * 兼容性   (Platform)   : CODESYS 3.5+ / TwinCAT 3 / 汇川 InoProShop / 施耐德 Machine Expert
 *                         仅依赖 Standard.library（ABS），零厂商私有库
 * 功能描述 (Function)   : 稳态偏置自适应修调（外挂修调器）：对闭环残差做带外积分、带内泄漏
 *                           |fErr| > fBand  →  _fTrim += fKiTrim × fErr × fCycle
 *                           |fErr| <= fBand →  _fTrim -= fLeak × _fTrim × fCycle
 *                         输出钳 [fTrimMin, fTrimMax] 并置 bSatLim。适用换热器结垢、阀门
 *                         磨损等缓慢漂移型稳态偏差的轻量外挂修正，不动主回路 PID 整定。
 * 接口     (Interface)  : 输入 fErr 闭环残差（工程单位）、bInService 投用、fKiTrim 修调积分
 *                         增益（1/s）、fBand 误差死区（工程单位）、fLeak 带内泄漏系数（1/s）、
 *                         fTrimMin/fTrimMax 修调限幅（工程单位）、fCycle 扫描周期（s，<=0
 *                         时用缺省周期）、bReset 复位；输出 fTrim 修调量、bSatLim 触限、
 *                         bError 故障标志。
 * 边界     (Boundary)   : ① **属主边界（写死）：本件只出修调偏置量，不注入任何回路、不接管
 *                         主 PID 整定**；注入点由上层叠加到设定值或输出偏置端。
 *                         ② bInService=FALSE 冻结不遗忘（退出即保持 _fTrim，防重投扰动，
 *                         语义写死不得由调用方假设）；bSatLim 复位。
 *                         ③ 非有限 fErr 当拍跳过（保持当拍 _fTrim 不动，R245）。
 *                         ④ fCycle <= 0 拒算，改用缺省扫描周期常量（防零周期积分跳变）。
 *                         ⑤ Anti-Windup：钳位后积分方向不改——限幅结果直接覆写 _fTrim，
 *                         不允许越限累积（`FB_DL_AntiWindupLink` 同族语义）。
 *                         ⑥ 组态闸：fTrimMin >= fTrimMax、fBand < 0、fLeak < 0 → 锁存
 *                         bError，冻结输出 fTrim=0 安全侧，解除沿 = bReset 上升沿。
 *                         ⑦ 零全局耦合（无 GVL / 无 VAR_EXTERNAL / 无物理地址）。
 * 分工声明 (Scope)      : 与 `FB_DL_Integrator` 分工：纯积分器无死区/泄漏/限幅闭环语义，
 *                         本件是带遗忘的闭环偏置修调；二者不互调不复制。
 * 来源标签 (Source Tag) : 自研线（带泄漏积分 clean-room）
 * 码表     (Codes)      : 本件不占用任何全局数字码位。出口为 LREAL 修调量 + BOOL 组；
 *                         数字码位待主控收口阶段统一派号。
 * 红线自检 (Redline)    : R1 ✓ 零 GVL/VAR_EXTERNAL ｜ R2 ✓ 零 %I/%Q/%M ｜ R3 ✓ 纯 IEC 61131-3
 *                         R4 ✓ 周期缺省闸 + 非有限跳过 + 钳位 Anti-Windup ｜ R5 ✓ 声明逐行同行双语注释
 *                         R6 N/A（无 ENUM 状态机） ｜ R7 ✓ 一 R_TRIG 段 0 无条件刷新
 * 修订历史 (Revision)   : 2026-11-20  v1.0.0  R48 首版（批次 2 · 序号 7）
 *                         验收向量：带外正残差积分上行；进入死区泄漏回落；触限后不累积；
 *                         退出投用冻结不遗忘；fCycle=0 用缺省周期。
 *==============================================================================*)

FUNCTION_BLOCK FB_DL_BiasAdaptiveTrim
VAR_INPUT
    fErr      : LREAL := 0.0;    // 闭环残差（被修调量实测与目标差） [工程单位] / Closed-loop residual
    bInService: BOOL := FALSE;   // 投用开关（FALSE=冻结保持不遗忘） [-] / In-service switch, FALSE freezes and holds
    fKiTrim   : LREAL := 0.1;    // 修调积分增益 [1/s] / Trim integral gain [1/s]
    fBand     : LREAL := 0.0;    // 误差死区半宽（带内不积分只泄漏） [工程单位] / Error deadband half-width
    fLeak     : LREAL := 0.0;    // 带内泄漏系数（遗忘速率） [1/s] / In-band leakage coefficient [1/s]
    fTrimMin  : LREAL := -10.0;  // 修调下限 [工程单位] / Trim lower limit
    fTrimMax  : LREAL := 10.0;   // 修调上限 [工程单位] / Trim upper limit
    fCycle    : LREAL := 0.0;    // 扫描周期（<=0 时用缺省周期） [s] / Scan cycle time, default used when <= 0
    bReset    : BOOL := FALSE;   // 复位，上升沿清组态故障锁存 [-] / Reset, rising edge clears config fault
END_VAR
VAR_OUTPUT
    fTrim   : LREAL;             // 修调偏置输出（已限幅） [工程单位] / Trim bias output, limited
    bSatLim : BOOL;              // 修调量触限（饱和发生，非故障） [-] / Trim hit the limit
    bError  : BOOL;              // 组态故障标志（锁存） [-] / Configuration fault flag, latched
END_VAR
VAR
    _fTrim    : LREAL := 0.0;    // 修调量锁存（投用退出即保持） / Latched trim, held when out of service
    _fCy      : LREAL;           // 当拍有效周期 [s] / Effective cycle this scan [s]
    _bErrLatch: BOOL;            // 组态故障锁存位（解除沿 = bReset 上升沿） / Latched config fault, cleared by reset edge
    rtReset   : R_TRIG;          // 复位沿实例，段 0 无条件调用 / Reset edge instance
    _bNonFin  : BOOL;            // 残差非有限当拍量 [-] / Non-finite residual this scan
    _fRaw     : LREAL;           // 当拍未限幅修调量 [工程单位] / Unlimited trim this scan
    _bSat     : BOOL;            // 当拍触限内部量（统一出口映射） / Saturation internal this scan
END_VAR
VAR CONSTANT
    DL_BAT_EPS      : LREAL := 1.0E-6;   // 浮点判零容差 [工程单位] / Float zero epsilon
    DL_BAT_CYCLEDEF : LREAL := 0.01;     // 缺省扫描周期（fCycle<=0 时启用） [s] / Default cycle time
    DL_BAT_ONE      : LREAL := 1.0;      // 单位常量（泄漏基） [无量纲] / Unit constant for leakage base
END_VAR

(* —— 段 0：非有限判 + 组态闸 + 周期派生 + 沿刷新 —— *)
_bNonFin := (fErr <> fErr) OR ((fErr - fErr) <> 0.0);       // 残差非有限（NaN 自不等 / Inf 差非零，R245） / Non-finite residual tests
IF (fTrimMin >= fTrimMax) OR (fBand < 0.0) OR (fLeak < 0.0) THEN
    _bErrLatch := TRUE;                                     // 组态域闸：锁存（R188 解除沿 = bReset 上升沿） / Config gate: latch
END_IF
IF fCycle > 0.0 THEN
    _fCy := fCycle;                                         // 组态周期有效 / Configured cycle valid
ELSE
    _fCy := DL_BAT_CYCLEDEF;                                // 周期缺省兜底（拒算零周期） / Default cycle fallback
END_IF
rtReset(CLK := bReset);                                     // 复位沿，每拍必调 / Reset edge, every scan

(* —— 段 1：复位沿 —— *)
IF rtReset.Q THEN
    _bErrLatch := FALSE;                                    // 清组态故障锁存 / Clear config fault latch
END_IF

(* —— 段 2：修调主算（未投用冻结不遗忘；故障期强制安全侧） —— *)
_bSat := FALSE;                                             // 触限内部量预清 / Saturation internal preset
IF _bErrLatch THEN
    _fTrim := 0.0;                                          // 故障安全侧：修调归零 / Fault safe side: trim forced zero
ELSIF NOT bInService THEN
    (* 未投用：_fTrim 冻结保持（防重投扰动，头注释②声明），bSatLim 复位 *)
    ;                                                       // 冻结分支无赋值（保持即语义） / Freeze branch holds by design
ELSIF _bNonFin THEN
    (* 残差非有限：当拍跳过积分与泄漏（保持 _fTrim 不动，R245） *)
    ;                                                       // 跳过分支保持 / Skip branch holds
ELSE
    IF ABS(fErr) > fBand THEN
        _fRaw := _fTrim + fKiTrim * fErr * _fCy;            // 带外积分：增益×残差×周期 / Out-of-band integration
    ELSE
        _fRaw := _fTrim - fLeak * _fTrim * _fCy;            // 带内泄漏：遗忘速率×修调×周期 / In-band leakage decay
    END_IF
    IF _fRaw > fTrimMax THEN
        _fTrim := fTrimMax;                                 // 上限覆写（Anti-Windup：不越限累积） / Ceiling overwrite, no windup
        _bSat := TRUE;                                      // 记触限 / Mark saturation
    ELSIF _fRaw < fTrimMin THEN
        _fTrim := fTrimMin;                                 // 下限覆写 / Floor overwrite
        _bSat := TRUE;                                      // 记触限 / Mark saturation
    ELSE
        _fTrim := _fRaw;                                    // 域内正常接受 / In-domain accept
    END_IF
END_IF

(* —— 段 3：出口单点映射（名实双出口同源，R191） —— *)
fTrim   := _fTrim;                                          // 修调量出口 / Trim outlet
bSatLim := _bSat AND (NOT _bErrLatch) AND bInService;       // 触限出口（冻结/故障期不复位不误报） / Saturation outlet
bError  := _bErrLatch;                                      // 故障标志出口 / Error flag outlet

END_FUNCTION_BLOCK

(* ---- FB_DL_BiquadCascade.st ---- *)
(*
  ==================================================================
  组件名 Component  : FB_DL_BiquadCascade
  分类   Category   : DL_Algo
  前缀   Naming     : FB_DL_ ｜ b/n/u/f/t/e/st 类型前缀制（R265）
  码位   Code ID    : 16#0002_3743 / 3744 / 3745 / 3748（故障级）
                      16#0002_3746 / 3747（信息级）
  版本   Version    : 1.0.0
  复杂度 Complexity  : 高
  功能   Purpose    : 多节二阶 IIR 级联（≤ 4 节，Direct Form II 每节独立状态），
                      用于高阶滤波（8 阶 = 4 节）现场组合；逐节 Jury 稳定闸。
  开源溯源 Origin    : 公开公式 clean-room，参考公开 DSP 教科书的二阶节级联结构与
                      Jury 稳定判据（分类与公式借鉴，零代码复制），本件实现、闸门
                      与码位 100% 自有。
  许可证 License    : MIT
  参考   Reference  : IEC 61131-3:2013 §6.6 算术运算符；Jury 三条件 |a2|<1 ∧
                      1+a1+a2>0 ∧ 1−a1+a2>0（与返修件 FB_DL_BiquadFilter v1.0.1
                      同源固化判据）
  平台   Platform   : 纯 IEC 61131-3（FOR / CASE / 四则 / ABS / R_TRIG），三平台通用
  依赖   Depends    : 仅 Standard.library（R_TRIG 属标准边沿检测）
  分工声明 Split     : FB_DL_BiquadFilter 为单节属主（R63 返修件，Jury 判据同源）；
                      本件多节级联，单节需求禁用本件（状态开销 ×4）；互引并注明
                      选型对照见 MANUAL_DL_Algo（R216）。
  归属 Ownership     : 本件无 TYPE 声明；全部引脚为 IEC 标准原生类型。
  ------------------------------------------------------------------
  边界 Boundary     :
                      一 逐节 Jury 稳定闸（返修 R2 固化判据）：任一**活动节**
                         （i < nStages）NOT (ABS(a2)<1 AND (1+a1+a2)>0 AND
                         (1−a1+a2)>0) → bCfgBad + 故障级 3744 + 三件套 + RETURN
                         结构早退（fOut 冻结最后有效值）；未激活节（i >= nStages）
                         的系数**不参与判据**（死节坏系数不误锁，写死）；
                      二 活动节系数任一非有限 → 故障级 3745（与 Jury 越域分码，
                         处置人不同：数值平台 / 算法工程师，R90）；
                      三 nStages 越域（< 1 或 > 4）或钳位域非法（fOutMin > fOutMax
                         或限值非有限）→ 故障级 3743（两组态场景出口同形：冻结 +
                         bCfgBad，R90 不另立）；
                      四 系数变更沿（任一活动系数 |新 − 旧| > 1.0E-9）→ 全链状态
                         清零（防新旧系数混算，BiquadFilter 同口径）+ 信息级 3747；
                      五 输出钳位 + bSat + 末活动节 w1 抗 windup 回写；非有限复检
                         → 故障级 3748 + 全链状态清零；
                      六 bEnable = FALSE 的语义写死（FB33-4 声明行）：fOut := 0 +
                         全链状态清零 + bValid = FALSE（下游控制量失能须归零）；
                      七 故障码锁存至 bResetState 上升沿回放（FB33-1 / R152）；
                         信息级逐拍重算不锁存；
                      八 段 0 无条件刷新 R_TRIG；CASE 无（线性级联，R6 标注 N/A）；
                         首拍 _bInit 全量初始化；无全局、无外部变量、无物理地址。
  错误码 Codes      :
    16#0002_3743【故障级】组态非法（nStages 越域 / 钳位域反序 / 限值非有限），锁存
    16#0002_3744【故障级】活动节系数越过 Jury 三条件稳定域，锁存
    16#0002_3745【故障级】活动节系数非有限（NaN 或 ±Inf），锁存
    16#0002_3748【故障级】输入 / 中间量 / 输出非有限（NaN 或 ±Inf），锁存
    16#0002_3746【信息级】本拍输出被钳位（bSat = TRUE，不锁存）
    16#0002_3747【信息级】系数变更沿触发全链状态清零（不锁存）
  码位反证 Note     :
    3743 / 3744 / 3745 / 3748 四码不可合并：四者的 bCfgBad 与 bValid 组合完全相同，
    但处置人不同（组态工程师 / 算法工程师 / 数值平台 / 现场仪表），仅靠输出组合无法
    还原成因，按 R90 分立（R90 反证句与返修件 FB_DL_BiquadFilter 同口径）。
  验收 Acceptance   :
    算法已证（脚本）：未跑 ｜ 编译器已证（三平台）：未跑
    V1 4 节低通级联（每节 RBJ 巴特沃斯 2 阶）阶跃 → 单调收敛无发散
    V2 节 3 系数失稳（a2 = −1.5, a1 = −1.9 违 Jury）→ bCfgBad + 全链冻结 + 3744
    V3 nStages = 0 / = 5 → 越域故障早退（3743）
    V4 节 4 系数坏但 nStages = 2 → 不影响（死节豁免，边界一回归向量）
    V5 在线改节 1 系数 → 全链清零 + 3747
    V6 bEnable = FALSE → fOut = 0、全链状态零、bValid = FALSE
    V7 输出大信号钳位 + bSat + 3746
  修订记录 Revision  :
    2026-11-21  v1.0.0  R63 首版（批 3 · 序号 8）
  ==================================================================
*)
FUNCTION_BLOCK FB_DL_BiquadCascade
VAR_INPUT
    bEnable     : BOOL := TRUE;    // 使能；FALSE 时输出归零并清全链状态（边界六）/ the enable, false zeroes the output and clears the chain
    bResetState : BOOL := FALSE;   // 状态复位电平，上升沿清全链状态与故障锁存 / the state reset level, its rising edge clears the chain and the fault latch
    fIn         : LREAL := 0.0;    // 输入量 [工程单位]，必须有限 / the input value, must be finite
    aB0         : ARRAY[0..3] OF LREAL; // 各节归一化前向系数 b0 [−] / the per stage normalized b0
    aB1         : ARRAY[0..3] OF LREAL; // 各节归一化前向系数 b1 [−] / the per stage normalized b1
    aB2         : ARRAY[0..3] OF LREAL; // 各节归一化前向系数 b2 [−] / the per stage normalized b2
    aA1         : ARRAY[0..3] OF LREAL; // 各节归一化反馈系数 a1 [−] / the per stage normalized a1
    aA2         : ARRAY[0..3] OF LREAL; // 各节归一化反馈系数 a2 [−] / the per stage normalized a2
    nStages     : DINT := 2;       // 节数 [节]，合法域 1..4 / the stage count, legal one to four
    fOutMin     : LREAL := -1.0E6; // 输出钳位域下界 [工程单位] / the output clamp floor
    fOutMax     : LREAL := 1.0E6;  // 输出钳位域上界 [工程单位] / the output clamp ceiling
END_VAR
VAR_OUTPUT
    fOut    : LREAL := 0.0;           // 滤波输出 [工程单位] / the filtered output
    bSat    : BOOL := FALSE;          // 本拍输出被钳位 [-] / the output was clamped on this scan
    bCfgBad : BOOL := FALSE;          // 组态非法（与故障锁存同源，锁存型）[-] / an illegal configuration latched with the fault
    bValid  : BOOL := FALSE;          // 输出可用 [-] / the output is usable
    eErr    : UDINT := 16#0000_0000;  // 错误码，0 = 正常 / the error code, zero is ok
    bError  : BOOL := FALSE;          // 故障锁存位（由锁存码派生，R99）/ the latched fault bit derived from the latched code
END_VAR
VAR
    _bInit   : BOOL := FALSE;                  // 首拍初始化标志（R310 / FB50-2）/ the first scan flag
    _afW1    : ARRAY[0..3] OF LREAL;           // 各节状态 w1 [工程单位] / the per stage state w1
    _afW2    : ARRAY[0..3] OF LREAL;           // 各节状态 w2 [工程单位] / the per stage state w2
    _afB0Prev : ARRAY[0..3] OF LREAL;          // 上拍 b0 快照 [−] / the previous b0 snapshots
    _afB1Prev : ARRAY[0..3] OF LREAL;          // 上拍 b1 快照 [−] / the previous b1 snapshots
    _afB2Prev : ARRAY[0..3] OF LREAL;          // 上拍 b2 快照 [−] / the previous b2 snapshots
    _afA1Prev : ARRAY[0..3] OF LREAL;          // 上拍 a1 快照 [−] / the previous a1 snapshots
    _afA2Prev : ARRAY[0..3] OF LREAL;          // 上拍 a2 快照 [−] / the previous a2 snapshots
    _fW      : LREAL := 0.0;                   // 本拍节内中间量 w [工程单位] / the intermediate w of this scan
    _fY      : LREAL := 0.0;                   // 本拍节内输出 y（级联传递量）[工程单位] / the stage output passed down the chain
    _fOutLast: LREAL := 0.0;                   // 最近一次有效输出（故障冻结源）[工程单位] / the last valid output used while frozen
    _nUse    : DINT := 0;                      // 钳位后的节数 [节] / the clamped stage count
    _i       : DINT := 0;                      // 节遍历索引 [下标] / the stage traversal index
    _iClr    : DINT := 0;                      // 清零遍历索引 [下标] / the clearing traversal index
    _bFinCoef: BOOL := FALSE;                  // 活动节系数有限闸结果（逐拍重算）/ the active stage finiteness gate result
    _bFinIn  : BOOL := FALSE;                  // 输入有限闸结果（逐拍重算）/ the input finiteness gate result
    _bFinDom : BOOL := FALSE;                  // 钳位限值有限闸结果（逐拍重算）/ the clamp limit finiteness gate result
    _bStable : BOOL := FALSE;                  // 活动节 Jury 闸结果（逐拍重算）/ the active stage Jury gate result
    _bCfgBadI: BOOL := FALSE;                  // 本拍组态非法标记（逐拍重算）/ the per scan configuration fault flag
    _bCoefChg: BOOL := FALSE;                  // 系数变更沿标记（逐拍重算，信息级 3747）/ the coefficient change flag
    _bSatI   : BOOL := FALSE;                  // 本拍钳位内部位 / the internal clamp bit
    _uLatch  : UDINT := 16#0000_0000;          // 故障码锁存（仅复位沿清除，FB33-1）/ the latched fault code cleared only by the reset edge
    rtReset  : R_TRIG;                         // 复位沿实例，段 0 无条件刷新（R7）/ the reset edge instance refreshed unconditionally
END_VAR  // R64 结构补齐：VAR 段缺失的 END_VAR（门禁机械修复）
VAR CONSTANT
    DL_BC_EPS   : LREAL := 1.0E-9;  // 系数变更判定容差 [−] / the coefficient change tolerance
    DL_BC_SMIN  : DINT := 1;        // 节数下界 [节] / the stage floor
    DL_BC_SMAX  : DINT := 4;        // 节数上界 [节] / the stage ceiling
    DL_BC_A2LIM : LREAL := 1.0;     // Jury 条件一 |a2| 边界 [−] / the Jury first condition boundary
    DL_BC_ONE   : LREAL := 1.0;     // Jury 条件二三的一常量 [−] / the unit constant of the Jury conditions
    DL_BC_ZERO  : LREAL := 0.0;     // 实数零常量 [工程单位] / the real zero constant
    DL_BC_ZEROI : DINT := 0;        // 整型零常量 [节] / the integer zero constant
    DL_BC_ONEI  : DINT := 1;        // 整型一常量 [节] / the integer one constant
END_VAR

// 段 0｜沿检测无条件周期刷新（禁入分支，R7）/ segment 0, the unconditional edge refresh
rtReset(CLK := bResetState); // 复位沿 / the reset edge

// 段 1｜首拍初始化（R310 / FB50-2；_bInit 与复位沿同款初始化）/ segment 1, the first scan init
IF NOT _bInit THEN // 首拍一拍 / the first scan
    _bInit := TRUE; // 置首拍标志 / raise the first scan flag
    FOR _iClr := DL_BC_ZEROI TO DL_BC_SMAX - DL_BC_ONE DO // 有界遍历全部节槽 / the bounded traversal over every stage slot
        _afW1[_iClr] := DL_BC_ZERO; // 状态 w1 显式清零 / clear the state w1 explicitly
        _afW2[_iClr] := DL_BC_ZERO; // 状态 w2 显式清零 / clear the state w2 explicitly
        _afB0Prev[_iClr] := aB0[_iClr]; // 系数快照对齐首拍值（防首拍误报变更沿）/ align the snapshot to avoid a spurious change edge
        _afB1Prev[_iClr] := aB1[_iClr]; // 快照对齐 / align the snapshot
        _afB2Prev[_iClr] := aB2[_iClr]; // 快照对齐 / align the snapshot
        _afA1Prev[_iClr] := aA1[_iClr]; // 快照对齐 / align the snapshot
        _afA2Prev[_iClr] := aA2[_iClr]; // 快照对齐 / align the snapshot
    END_FOR
    _fOutLast := DL_BC_ZERO; // 最近有效输出显式清零 / clear the last valid output explicitly
    _uLatch := 16#0000_0000; // 故障码锁存显式清零 / clear the latched code explicitly
END_IF
IF rtReset.Q THEN // 复位沿（作用域：清锁存 + 清全链状态，R311 声明）/ the reset edge with the declared scope
    _uLatch := 16#0000_0000; // 清故障码锁存（唯一的故障解除路径）/ clear the latched code, the only release path
    FOR _iClr := DL_BC_ZEROI TO DL_BC_SMAX - DL_BC_ONE DO // 有界遍历全部节槽 / the bounded traversal over every stage slot
        _afW1[_iClr] := DL_BC_ZERO; // 清状态 w1 / clear the state w1
        _afW2[_iClr] := DL_BC_ZERO; // 清状态 w2 / clear the state w2
    END_FOR
END_IF
_bSatI := FALSE; // 钳位单拍内部位预清零 / preset the internal clamp bit false
_bCoefChg := FALSE; // 系数变更标记预清零 / preset the coefficient change flag false
_bCfgBadI := FALSE; // 组态非法标记预清零 / preset the configuration fault flag false

// 段 2｜组态闸（边界一三：nStages 越域 / 钳位域 / 活动节系数非有限 / Jury，成因独立码 R190）/ segment 2, the configuration gates
_nUse := nStages; // 节数接管 [节] / take the stage count
IF (_nUse < DL_BC_SMIN) OR (_nUse > DL_BC_SMAX) THEN // 节数越域 / the stage count is out of the domain
    _bCfgBadI := TRUE; // 置组态标记 / raise the configuration flag
    IF _uLatch = 16#0000_0000 THEN // 仅首因入锁存（R152）/ latch only the first cause
        _uLatch := 16#0002_3743; // 故障级：组态非法（节数越域）/ fault grade, an illegal configuration
    END_IF
    IF _nUse < DL_BC_SMIN THEN // 下界钳位（防遍历越界）/ the floor clamp for the traversal safety
        _nUse := DL_BC_SMIN; // 钳到一节 / clamp to one stage
    ELSE // 上界钳位 / the ceiling clamp
        _nUse := DL_BC_SMAX; // 钳到四节 / clamp to four stages
    END_IF
END_IF
_bFinDom := (fOutMin = fOutMin) AND ((fOutMin - fOutMin) = (fOutMin - fOutMin))
         AND (fOutMax = fOutMax) AND ((fOutMax - fOutMax) = (fOutMax - fOutMax)); // 限值有限 / the limits are finite
IF (NOT _bFinDom) OR (fOutMin > fOutMax) THEN // 限值非有限或域反序 / the limits are not finite or the domain is reversed
    _bCfgBadI := TRUE; // 置组态标记 / raise the configuration flag
    IF _uLatch = 16#0000_0000 THEN // 仅首因入锁存 / latch only the first cause
        _uLatch := 16#0002_3743; // 故障级：组态非法（钳位域）/ fault grade, an illegal clamp domain
    END_IF
END_IF
_bFinIn := (fIn = fIn) AND ((fIn - fIn) = (fIn - fIn)); // 输入有限 / the input is finite
FOR _i := DL_BC_ZEROI TO _nUse - DL_BC_ONE DO // 有界遍历活动节（死节豁免，边界一）/ the bounded traversal over the active stages, dead stages exempt
    _bFinCoef := (aB0[_i] = aB0[_i]) AND ((aB0[_i] - aB0[_i]) = (aB0[_i] - aB0[_i]))
              AND (aB1[_i] = aB1[_i]) AND ((aB1[_i] - aB1[_i]) = (aB1[_i] - aB1[_i]))
              AND (aB2[_i] = aB2[_i]) AND ((aB2[_i] - aB2[_i]) = (aB2[_i] - aB2[_i]))
              AND (aA1[_i] = aA1[_i]) AND ((aA1[_i] - aA1[_i]) = (aA1[_i] - aA1[_i]))
              AND (aA2[_i] = aA2[_i]) AND ((aA2[_i] - aA2[_i]) = (aA2[_i] - aA2[_i])); // 本节五系数有限 / the five coefficients of this stage are finite
    _bStable := (ABS(aA2[_i]) < DL_BC_A2LIM) AND ((DL_BC_ONE + aA1[_i] + aA2[_i]) > DL_BC_ZERO) AND ((DL_BC_ONE - aA1[_i] + aA2[_i]) > DL_BC_ZERO); // Jury 三条件（与 FB_DL_BiquadFilter v1.0.1 同口径）/ the Jury three conditions aligned with the single stage owner
    IF (NOT _bFinCoef) AND (_uLatch = 16#0000_0000) THEN // 成因：活动节系数非有限（不覆盖已有首因）/ the coefficients of an active stage are not finite
        _bCfgBadI := TRUE; // 置组态标记 / raise the configuration flag
        _uLatch := 16#0002_3745; // 故障级：活动节系数非有限 / fault grade, the coefficients are not finite
        bError := TRUE; // 同拍置故障标志（R45 配对，段 4 故障分支沿用）/ raise the fault flag on the same scan
    ELSIF (NOT _bStable) AND (_uLatch = 16#0000_0000) THEN // 成因：活动节越 Jury 域 / the Jury conditions are exceeded
        _bCfgBadI := TRUE; // 置组态标记 / raise the configuration flag
        _uLatch := 16#0002_3744; // 故障级：活动节越过 Jury 三条件稳定域 / fault grade, the Jury conditions are exceeded
        bError := TRUE; // 同拍置故障标志（R45 配对，段 4 故障分支沿用）/ raise the fault flag on the same scan
    END_IF
END_FOR
IF (NOT _bFinIn) AND (_uLatch = 16#0000_0000) THEN // 成因：输入非有限（不覆盖已有首因）/ the input is not finite
    _uLatch := 16#0002_3748; // 故障级：输入非有限 / fault grade, the input is not finite
END_IF

// 段 3｜使能失能分支最先消费：降级为安全值并清全链（边界六声明行）/ segment 3, the disabled branch degrades to the safe value
IF NOT bEnable THEN // 失能 / disabled
    FOR _iClr := DL_BC_ZEROI TO DL_BC_SMAX - DL_BC_ONE DO // 有界遍历全部节槽 / the bounded traversal over every stage slot
        _afW1[_iClr] := DL_BC_ZERO; // 状态清零（失能即弃用历史）/ clear the state, the history is abandoned
        _afW2[_iClr] := DL_BC_ZERO; // 状态清零 / clear the state
    END_FOR
    _fOutLast := DL_BC_ZERO; // 输出归零（下游控制量失能须归零，非冻结末值）/ zero the output, a control quantity must fall to zero
    fOut := DL_BC_ZERO; // 出口归零 [工程单位] / the outlet falls to zero
    bSat := FALSE; // 钳位位清零 / clear the clamp bit
    bCfgBad := (_uLatch <> 16#0000_0000); // 组态标记照实回放（与锁存同源）/ replay the configuration flag from the latch
    bValid := FALSE; // 输出不可用（安全值不是滤波结果，明示而非静默）/ mark the output unusable, a safe zero is not a filter result
    bError := (_uLatch <> 16#0000_0000); // 故障位照实回放 / replay the fault bit from the latch
    eErr := _uLatch; // 故障码锁存回放（信息级不参与失能分支）/ replay the latched code
    RETURN; // 早退，不推进级联 / early return without advancing the chain
END_IF

// 段 4｜组态故障：冻结最近有效输出，不推进状态（边界一五，结构早退；冻结源做有限性闸，FB51-3）/ segment 4, freeze on a fault without advancing the chain
IF (_uLatch <> 16#0000_0000) OR _bCfgBadI THEN // 任一故障相 / any fault phase
    IF (_fOutLast = _fOutLast) AND ((_fOutLast - _fOutLast) = (_fOutLast - _fOutLast)) THEN // 冻结源有限性闸（冻结只防推进不防污染）/ the frozen source finiteness gate
        fOut := _fOutLast; // 冻结最近有效输出 [工程单位] / freeze the last valid output
    ELSE // 冻结源自身被污染（理论上不可达）/ the frozen source itself is polluted
        _fOutLast := DL_BC_ZERO; // 归零重建 / rebuild from zero
        fOut := DL_BC_ZERO; // 出口归零 [工程单位] / the outlet falls to zero
    END_IF
    bSat := FALSE; // 钳位位清零 / clear the clamp bit
    bCfgBad := _bCfgBadI OR (_uLatch = 16#0002_3743) OR (_uLatch = 16#0002_3744) OR (_uLatch = 16#0002_3745); // bCfgBad 专指组态族三码，3748 输入坏不复用 / the configuration flag covers only the configuration family codes
    bValid := FALSE; // 输出不可用 / the output is not usable
    bError := TRUE; // 故障位置位 / raise the fault bit
    eErr := _uLatch; // 锁存码回放（不按当下输入重新推断，R152）/ replay the latched code
    RETURN; // 结构早退 / the structural early exit
END_IF

// 段 5｜系数变更沿：任一活动系数 |新 − 旧| > 容差即清全链状态（边界四）/ segment 5, the coefficient change edge clears the chain
FOR _i := DL_BC_ZEROI TO _nUse - DL_BC_ONE DO // 有界遍历活动节 / the bounded traversal over the active stages
    IF (ABS(aB0[_i] - _afB0Prev[_i]) > DL_BC_EPS) OR (ABS(aB1[_i] - _afB1Prev[_i]) > DL_BC_EPS)
    OR (ABS(aB2[_i] - _afB2Prev[_i]) > DL_BC_EPS) OR (ABS(aA1[_i] - _afA1Prev[_i]) > DL_BC_EPS)
    OR (ABS(aA2[_i] - _afA2Prev[_i]) > DL_BC_EPS) THEN // 本节任一系数变更 / any coefficient of this stage changed
        _bCoefChg := TRUE; // 置变更标记（信息级 3747）/ raise the change flag
        FOR _iClr := DL_BC_ZEROI TO DL_BC_SMAX - DL_BC_ONE DO // 有界遍历全部节槽（全链清零防混算）/ the bounded traversal over every slot
            _afW1[_iClr] := DL_BC_ZERO; // 清状态 w1 / clear the state w1
            _afW2[_iClr] := DL_BC_ZERO; // 清状态 w2 / clear the state w2
        END_FOR
    END_IF
    _afB0Prev[_i] := aB0[_i]; // 系数快照推进 [−] / advance the b0 snapshot
    _afB1Prev[_i] := aB1[_i]; // 快照推进 [−] / advance the b1 snapshot
    _afB2Prev[_i] := aB2[_i]; // 快照推进 [−] / advance the b2 snapshot
    _afA1Prev[_i] := aA1[_i]; // 快照推进 [−] / advance the a1 snapshot
    _afA2Prev[_i] := aA2[_i]; // 快照推进 [−] / advance the a2 snapshot
END_FOR

// 段 6｜逐节 Direct Form II 递推（节间串接：本拍节输出即下一节输入）/ segment 6, the per stage recursion chained down
_fY := fIn; // 级联入口 = 输入 [工程单位] / the chain inlet is the input
FOR _i := DL_BC_ZEROI TO _nUse - DL_BC_ONE DO // 有界遍历活动节 / the bounded traversal over the active stages
    _fW := _fY - (aA1[_i] * _afW1[_i]) - (aA2[_i] * _afW2[_i]); // 节内中间量 w [工程单位] / the intermediate w of this stage
    _fY := (aB0[_i] * _fW) + (aB1[_i] * _afW1[_i]) + (aB2[_i] * _afW2[_i]); // 节输出 y [工程单位] / the stage output
    _afW2[_i] := _afW1[_i]; // 状态右移：w1 → w2 / shift the state
    _afW1[_i] := _fW; // 状态推进：本拍 w → w1 / advance the state
END_FOR

// 段 7｜输出钳位 + 末活动节 w1 抗 windup 状态回写 / segment 7, the clamp with the anti windup write back
IF _fY > fOutMax THEN // 超上界 / above the ceiling
    fOut := fOutMax; // 钳上界 [工程单位] / clamp to the ceiling
    _bSatI := TRUE; // 置钳位内部位 / raise the internal clamp bit
    _afW1[_nUse - DL_BC_ONE] := fOutMax; // 末活动节状态回写（防积分式累积发散）[工程单位] / write the last active state back
ELSIF _fY < fOutMin THEN // 超下界 / below the floor
    fOut := fOutMin; // 钳下界 [工程单位] / clamp to the floor
    _bSatI := TRUE; // 置钳位内部位 / raise the internal clamp bit
    _afW1[_nUse - DL_BC_ONE] := fOutMin; // 末活动节状态回写 [工程单位] / write the state back
ELSE // 域内 / inside the domain
    fOut := _fY; // 直出输出 [工程单位] / pass the output through
END_IF

// 段 8｜全部内部量非有限复检：污染即拒收并锁存（FB32-7 保持槽口径）/ segment 8, the finiteness recheck before the states are stored
IF (fOut <> fOut) OR ((fOut - fOut) <> (fOut - fOut))
OR (_fY <> _fY) OR ((_fY - _fY) <> (_fY - _fY)) THEN // 输出或级联传递量非有限（NaN 自反 / Inf 差值自减）/ a non finite output or intermediate
    FOR _iClr := DL_BC_ZEROI TO DL_BC_SMAX - DL_BC_ONE DO // 有界遍历全部节槽 / the bounded traversal over every slot
        _afW1[_iClr] := DL_BC_ZERO; // 状态清零，禁污染物驻留 / clear the state so nothing polluted remains
        _afW2[_iClr] := DL_BC_ZERO; // 状态清零 / clear the state
    END_FOR
    IF _uLatch = 16#0000_0000 THEN // 仅首因入锁存 / latch only the first cause
        _uLatch := 16#0002_3748; // 故障级：输入或中间量非有限 / fault grade, the input or the intermediate is not finite
    END_IF
    fOut := DL_BC_ZERO; // 出口归零 [工程单位] / the outlet falls to zero
    bSat := FALSE; // 钳位位清零 / clear the clamp bit
    bCfgBad := FALSE; // 3748 属测量坏而非组态坏 / the input fault is a measurement issue
    bValid := FALSE; // 输出不可用 / the output is not usable
    bError := TRUE; // 故障位置位 / raise the fault bit
    eErr := _uLatch; // 锁存码回放 / replay the latched code
    RETURN; // 早退 / early return
END_IF

// 段 9｜最近有效输出写回（写前已过非有限闸）/ segment 9, store the last valid output
_fOutLast := fOut; // 快照更新 [工程单位] / update the snapshot

// 段 10｜统一出口（单拍位映射 + 信息级重算，R187 / FB51-8）/ segment 10, the unified outlet
bSat := _bSatI; // 钳位位出口 / the clamp bit outlet
bCfgBad := (_uLatch = 16#0002_3743) OR (_uLatch = 16#0002_3744) OR (_uLatch = 16#0002_3745); // 组态标记出口（与锁存同源，3748 不复用）/ the configuration flag outlet from the latch
bValid := TRUE; // 域内输出可用 / the in-domain output is usable
bError := (_uLatch <> 16#0000_0000); // 故障位出口（锁存派生，R99）/ the fault bit outlet derived from the latch
IF _uLatch <> 16#0000_0000 THEN // 故障锁存回放优先 / the latched fault replays first
    eErr := _uLatch; // 锁存码 [码] / the latched code
ELSIF _bSatI THEN // 输出钳位（信息级，逐拍重算）/ the output clamp, informational
    eErr := 16#0002_3746; // 信息级：本拍输出被钳位 / informational, the output was clamped
ELSIF _bCoefChg THEN // 系数变更（信息级，逐拍重算）/ the coefficient change, informational
    eErr := 16#0002_3747; // 信息级：系数变更沿触发全链状态清零 / informational, a coefficient change cleared the chain
ELSE // 无事件 / no event
    eErr := 16#0000_0000; // 正常 / ok
END_IF
END_FUNCTION_BLOCK

(* ---- FB_DL_BumplessHandAuto.st ---- *)
(*
  组件名 Component   : FB_DL_BumplessHandAuto
  子库 Sublibrary    : DL_Algo
  版本 Version       : 1.0.0
  兼容性 Platform    : CODESYS 3.5 / TwinCAT 3 / 汇川 InoProShop / Machine Expert（仅 Standard.library）
  功能 Function      : 手/自动无扰切换（T0 标准语义件）：
                       1) 手动相：输出 = fManualOut，同时以自动需求做双向跟踪监督；
                       2) 切自动：切换偏差 |fAutoOut - 当前输出| <= fSwDevMaxPct 时直接无扰
                       切入；超限时经 eAutoRamp 相以 fSwRampPctS 斜率逼近自动需求后切入；
                       3) 切手动：输出立即跟随 fManualOut（跟踪量恒可用，无扰返回）；
                       4) 跟踪失效报警：手动相下执行器反馈偏离手动指令超 fTrackTolPct
                       持续 tTrackTo → 报警锁存（故障级，bReset 上升沿解除）。
  边界 Boundary      : ① 本件只做输出选择与切换监督，不内嵌 PID（需求由上层回路提供）；
                       ② 除法/斜率换算前置域闸：fSwRampPctS <= 0 判组态非法；
                       ③ 非有限值（NaN 自反 + 无穷差值自减）判输入非法，锁存安全侧；
                       ④ eAutoRamp 相退出双条件：偏差入容差（达成）或需求翻转回手动；
                       ⑤ 故障锁存解除唯一路径 = bReset 上升沿（输入引脚，恒可达）；
                       ⑥ 无全局变量引用、无外部变量声明、无物理地址寻址。
  依赖 Depends       : Standard.library（R_TRIG / TON）
  溯源 Origin        : IEC 61131-3 标准语义的道莅防御性实现（双向跟踪无扰切换为标准
                       控制回路手/自动语义，T0 口径）
  码位 Code          : 16#02_3_8B
  码表 Error codes（Algo 格 02_3_8B，单轨：故障 0x038B / 信息 0x028B）:
    16#0002_038B 故障级：跟踪失效锁存（手动相反馈偏离超容差持续 tTrackTo）或
                 组态非法/输入非有限，锁存至 bReset 上升沿
    16#0002_028B 信息级：斜坡切入自动沿（eAutoRamp → eAuto 迁移拍）
  修订历史 Revision  :
    2026-11-19  v1.0.0  R44 首版（批次 1 · 序号 4）
*)

TYPE E_DL_BhaState :
(
    eManual   := 0,    // 手动：输出跟随手动指令 / Manual, output follows hand command
    eAutoRamp := 10,   // 斜坡：输出限速逼近自动需求 / Ramp, output slews to auto demand
    eAuto     := 20,   // 自动：输出 = 自动需求 / Auto, output equals auto demand
    eFault    := 90    // 故障：跟踪失效或组态锁存 / Fault, latched
);
END_TYPE

FUNCTION_BLOCK FB_DL_BumplessHandAuto
VAR_INPUT
    bAutoMode   : BOOL;                    // 自动模式请求（电平）[-] / Auto mode request
    bReset      : BOOL;                    // 上升沿清故障锁存 [-] / Reset edge
    fAutoOut    : REAL;                    // 自动需求（上层回路输出）[%] / Auto demand
    fManualOut  : REAL;                    // 手动指令 [%] / Manual command
    fFbPos      : REAL;                    // 执行器反馈位置 [%] / Actuator feedback
    fSwDevMaxPct: REAL := 10.0;            // 直接切换允许偏差 [%] / Direct switch deviation limit
    fSwRampPctS : REAL := 20.0;            // 斜坡切入速率 [%/秒] / Switch slew rate
    fTrackTolPct: REAL := 5.0;             // 跟踪容差 [%] / Tracking tolerance
    tTrackTo    : TIME := T#5S;            // 跟踪失效确认窗 [毫秒] / Tracking fail confirm window
    tCycle      : TIME := T#10MS;          // 扫描周期 [毫秒] / Scan cycle time
END_VAR
VAR_OUTPUT
    fOut        : REAL;                    // 选择输出 [%] / Selected output
    bAuto       : BOOL;                    // 自动相电平标志 [-] / Auto state level
    bRamping    : BOOL;                    // 斜坡相电平标志 [-] / Ramping state level
    bError      : BOOL;                    // 故障锁存标志 [-] / Fault latch flag
    uErrId      : UDINT;                   // 事件码，0 = 无事件 / Event code
    eState      : E_DL_BhaState;           // 状态出口，段尾单点映射 / State outlet
END_VAR
VAR
    rtReset     : R_TRIG;                  // 复位沿实例，段 0 无条件刷新 / Reset edge
    rtToAuto    : R_TRIG;                  // 切自动沿实例，段 0 无条件刷新 / To-auto edge
    rtToManual  : R_TRIG;                  // 切手动沿实例，段 0 无条件刷新 / To-manual edge
    tonTrackTo  : TON;                     // 跟踪失效确认（专用超时件命名（R228A 豁免））/ Tracking timeout
    _eState     : E_DL_BhaState := E_DL_BhaState.eManual;   // 内部相位（CASE 唯一写入目标）/ Internal phase
    _fDev       : REAL;                    // 切换偏差绝对值 [%] / Switch deviation
    _fFbDev     : REAL;                    // 跟踪偏差绝对值 [%] / Tracking deviation
    _fStep      : REAL;                    // 本拍斜坡步长 [%] / Slew step per scan
    _fCyS       : REAL;                    // 扫描周期秒值 [秒] / Cycle seconds
    _bFault     : BOOL;                    // 故障锁存位（锁存量） / Latched fault bit
    _uFault     : UDINT;                   // 故障码锁存（锁存量） / Latched fault code
    _bCfgBad    : BOOL;                    // 组态非法当拍量 [-] / Config illegal flag
    _bNonFin    : BOOL;                    // 输入非有限当拍量 [-] / Non-finite input flag
END_VAR
VAR CONSTANT
    DL_DEV_EPS  : REAL := 1.0E-6;          // 偏差入容差判据 [％] / Deviation snap tolerance
    DL_ABS_MAX  : REAL := 1.0E30;          // 有限值判定上界 [%] / Finite value bound
    DL_ZERO     : REAL := 0.0;             // 零常量 [%] / Zero constant
    DL_MS_PER_S : REAL := 1000.0;          // 毫秒 → 秒换算系数 [毫秒/秒] / Milliseconds per second
END_VAR

(* —— 段 0｜沿与定时器每拍无条件刷新（禁置于 IF/CASE 内） —— *)
_fFbDev := ABS(fFbPos - fManualOut);     // 跟踪偏差先行计算，供定时器 IN 引用
rtReset   (CLK := bReset);
rtToAuto  (CLK := bAutoMode);
rtToManual(CLK := NOT bAutoMode);
tonTrackTo(IN := (_eState = E_DL_BhaState.eManual) AND (_fFbDev > fTrackTolPct) AND (NOT _bFault),
           PT := tTrackTo);

(* —— 段 1｜瞬时量预清零与周期换算（锁存量 _bFault/_uFault 不入清单） —— *)
uErrId   := 16#0000_0000;
_bCfgBad := FALSE;
_bNonFin := FALSE;
_fCyS    := TIME_TO_REAL(tCycle) / DL_MS_PER_S;

(* —— 段 2｜复位沿：故障一次性清干净，相位回手动（安全侧待机） —— *)
IF rtReset.Q THEN
    _bFault := FALSE;
    _uFault := 16#0000_0000;
    _eState := E_DL_BhaState.eManual;    // 复位后回手动待机，由沿重新切入自动
END_IF

(* —— 段 3｜组态闸与输入非有限判据 —— *)
IF (fSwRampPctS <= DL_ZERO) OR (fSwDevMaxPct < DL_ZERO) OR (fTrackTolPct <= DL_ZERO)
   OR (tCycle = T#0S) THEN
    _bCfgBad := TRUE;
END_IF
IF (fAutoOut <> fAutoOut) OR ((fAutoOut - fAutoOut) <> DL_ZERO)
   OR (fManualOut <> fManualOut) OR ((fManualOut - fManualOut) <> DL_ZERO)
   OR (fFbPos <> fFbPos) OR ((fFbPos - fFbPos) <> DL_ZERO) THEN
    _bNonFin := TRUE;
END_IF

(* —— 段 4｜故障触发：组态/输入非法或跟踪失效（tonTrackTo.Q 为保持量级判据） —— *)
IF _bCfgBad OR _bNonFin THEN
    _bFault := TRUE;
    _uFault := 16#0002_038B;
    _eState := E_DL_BhaState.eFault;
ELSIF (_eState = E_DL_BhaState.eManual) AND tonTrackTo.Q THEN
    _bFault := TRUE;                     // 手动相跟踪失效：反馈偏离超容差持续超窗
    _uFault := 16#0002_038B;
    _eState := E_DL_BhaState.eFault;
END_IF

(* —— 段 5｜主状态机：四态全覆盖 + ELSE 兜底 —— *)
CASE _eState OF

E_DL_BhaState.eManual:
    fOut   := fManualOut;                // 输出跟随手动指令
    bAuto  := FALSE;
    bRamping := FALSE;
    ;                                    // 跟踪监督判据 _fFbDev 已在段 0 预算，经 tonTrackTo 承载
    IF rtToAuto.Q AND (NOT _bFault) THEN
        _fDev := ABS(fAutoOut - fOut);
        IF _fDev <= fSwDevMaxPct THEN
            _eState := E_DL_BhaState.eAuto;      // 小偏差直接无扰切入
        ELSE
            _eState := E_DL_BhaState.eAutoRamp;  // 大偏差限速逼近
        END_IF
    END_IF

E_DL_BhaState.eAutoRamp:
    bAuto    := FALSE;
    bRamping := TRUE;
    _fStep   := fSwRampPctS * _fCyS;     // 本拍步长 = 速率 × 周期
    IF fOut < fAutoOut THEN
        fOut := MIN(fOut + _fStep, fAutoOut);    // 上行逼近，不越过需求
    ELSIF fOut > fAutoOut THEN
        fOut := MAX(fOut - _fStep, fAutoOut);    // 下行逼近，不越过需求
    END_IF
    IF ABS(fAutoOut - fOut) <= DL_DEV_EPS THEN
        uErrId  := 16#0002_028B;         // 信息级：斜坡切入自动沿
        _eState := E_DL_BhaState.eAuto;  // 迁出条件 1：偏差达成
    ELSIF rtToManual.Q THEN
        _eState := E_DL_BhaState.eManual;    // 迁出条件 2：需求翻转回手动
    END_IF

E_DL_BhaState.eAuto:
    fOut      := fAutoOut;               // 输出 = 自动需求
    bAuto     := TRUE;
    bRamping  := FALSE;
    IF rtToManual.Q THEN
        _eState := E_DL_BhaState.eManual;    // 无扰返回：手动相输出立即跟手
    END_IF

E_DL_BhaState.eFault:
    bError := TRUE;                      // 故障相驻留：出口冻结保持，只认复位沿（段 2 迁出）
    ;                                    // （故障相 fOut 保持最后值，禁止任何迁移）

ELSE
    _bFault := TRUE;                     // 兜底：非法相位锁存
    _uFault := 16#0002_038B;
    bError  := TRUE;
    _eState := E_DL_BhaState.eFault;
END_CASE

(* —— 段 6｜状态出口单点映射 —— *)
eState := _eState;
END_FUNCTION_BLOCK

(* ---- FB_DL_BumplessTransfer.st ---- *)
(*
    FB_DL_BumplessTransfer —— 手 / 自动无扰切换
    ------------------------------------------------------------------
    分类      : DL_Algo / Control
    前缀      : FB_DL_
    版本      : 1.0.0
    溯源      : T2-5 Mod_PID（源矩阵明列「参数域已取尽，后续仅剩手自动切换手册细节」，
                本件即该细节的收口件）；T1-1 OSCAT Basic 反作用增益惯例作次源对照；
                无扰过渡律、状态机、码位 100% 自有；clean-room 重写，未复制任何
                闭源厂商源码，参考实现仅限 MIT/Apache 许可
    平台      : 纯 IEC 61131-3，CODESYS V3.5+ / TwinCAT 3 / InoProShop 通用
    作者      : 道莅代码库 · PLC编程专家（R18）
    ------------------------------------------------------------------
    功能说明  : 手动到自动切换时，输出从「手动末值」按限斜率过渡到「PID 输出」，
                杜绝阀门 / 变频器被给定量阶跃冲击（水锤、皮带打滑、加热丝浪涌）；
                手动期持续把输出跟踪到实际反馈（反算跟踪），使自动接管时积分项不突跳；
                过渡收敛判据用「偏差不大于单拍步长加容差」，浮点判等全部带容差；
                输出限幅为双侧，只做单侧限幅是本库明令禁止的常见缺陷；
                职责边界：本件不内联 PID，PID 输出由上层注入，避免两套积分器打架。
    错误码    : 16#0002_2401 过渡中偏差超提示窗（正常现象，非故障）——信息级，不置故障
                16#0002_2402 预留禁用（信息级，不得挪用）
                16#0002_2410 斜率参数非法（不在 0.01~1000 %/s）——故障级，过渡禁用直接取 PID 输出
                16#0002_2411 给定非有限（NaN / 正负 INF）或状态机落 ELSE 兜底——故障级，保持末次输出
                16#0002_2412 预留禁用（故障级，不得挪用）
    码位总账  : 16#0002_2401 用 / 16#0002_2402 预留 ｜ 16#0002_2410 用 / 16#0002_2411 用 / 16#0002_2412 预留
    状态机    : E_DL_TransferState（eIdle / eManual / eTransfer / eAuto / eFault），
                CASE 含 ELSE 兜底，兜底固定置 eFault 与 2411
    采样约定  : fbTrigReset 在本体首部无条件刷新；单拍步长按固定任务周期常量
                DL_TR_DT 折算，必须与实际任务周期一致，周期改动须同步改该常量。
    修订记录  : 2026-11-16 v1.0.0 首次入库（R18）
*)

(*-----------------------------------------------------------------------------
 * 枚举: E_DL_TransferState（归属本功能块，与其同文件发布）
 * 含义: 手自动无扰切换状态机离散态，步长 10 留空位，故障态取 99 排末位
 *----------------------------------------------------------------------------*)
TYPE E_DL_TransferState :
(
    eIdle     := 0,    // 空闲：输出归零，等待首次使能 / Idle, output zeroed, waiting for the first enable
    eManual   := 10,   // 手动：输出跟踪实际反馈，为接管做准备 / Manual, output tracks the actual feedback to prepare the takeover
    eTransfer := 20,   // 过渡：按限斜率逼近 PID 输出 / Transfer, approaching the PID output at the limited rate
    eAuto     := 30,   // 自动：输出直接等于 PID 输出 / Auto, output equals the PID output
    eFault    := 99    // 故障锁存：给定非有限或非法状态，保持末次输出 / Fault latched, non-finite setpoint or illegal state, holds the last output
) UINT;
END_TYPE

FUNCTION_BLOCK FB_DL_BumplessTransfer
VAR_INPUT
    bEnable     : BOOL;                        // 使能，FALSE 输出 0 并清过渡 / enable, FALSE zeroes the output and clears the transfer
    bReset      : BOOL;                        // 复位，上升沿放弃过渡直接取目标值（调试用）/ reset, rising edge abandons the transfer and takes the target directly, commissioning only
    bAuto       : BOOL := FALSE;               // TRUE 自动 / FALSE 手动 / TRUE auto, FALSE manual
    fManualOut  : REAL := 0.0;                 // 手动给定，仅手动期生效 [%]，范围 -100.0~100.0 / manual setpoint, manual mode only [%], range -100.0~100.0
    fPidOut     : REAL := 0.0;                 // PID 输出，由上层注入，本件不内联 PID [%] / PID output injected by the caller, no PID inside [%]
    fTrackVal   : REAL := 0.0;                 // 手动期跟踪目标，一般接实际阀位反馈 [%]，范围 -100.0~100.0 / tracking target during manual mode, usually the actual valve position [%], range -100.0~100.0
    fRateMax    : REAL := 10.0;                // 过渡最大变化率 [%/s]，范围 0.01~1000.0 / maximum transfer rate [%/s], range 0.01~1000.0
    fDevWindow  : REAL := 5.0;                 // 过渡偏差提示窗 [%] / deviation hint window during the transfer [%]
END_VAR
VAR_OUTPUT
    fOut         : REAL;                       // 最终输出，双侧限幅 [%] / final output, clamped on both sides [%]
    bTracking    : BOOL;                       // 手动期跟踪中 / tracking during manual mode
    bInTransfer  : BOOL;                       // 自动接管过渡中 / transfer in progress
    fDeviation   : REAL;                       // 当前输出与 PID 输出的偏差 [%] / deviation between the output and the PID output [%]
    tInTransfer  : TIME;                       // 已过渡时长 [ms] / elapsed transfer time [ms]
    eErr         : UDINT;                      // 错误码，0=正常 / error id, 0=ok
    bError       : BOOL;                       // 故障标志，eErr 为故障级时 TRUE / error flag, TRUE on fault-level eErr
END_VAR
VAR
    fbTrigReset : R_TRIG;                      // 复位沿检测实例，本体首部无条件刷新 / reset edge instance, refreshed unconditionally
    eState      : E_DL_TransferState := E_DL_TransferState.eIdle; // 内部状态机步序 / internal state machine step
    fLastOut    : REAL;                        // 上一拍输出，过渡起点 [%] / previous cycle output, the transfer starting point [%]
    fStep       : REAL;                        // 单拍允许变化量 [%] / allowed change per cycle [%]
    tLast       : TIME;                        // 过渡累计时长 [ms] / accumulated transfer time [ms]
    tDelta      : TIME;                        // 本拍时间增量，取固定任务周期 [ms] / time increment of this cycle, the fixed task period [ms]
    bInit       : BOOL := FALSE;               // 首扫标志，初值 FALSE，判据 NOT bInit / first-scan flag, initial FALSE, tested with NOT
    bNonFin     : BOOL;                        // 给定非有限判定标志 / setpoint non-finite flag
    bRateOk     : BOOL;                        // 斜率参数合法标志 / rate parameter valid flag
    fClamped    : REAL;                        // 限幅中间量 [%] / clamping intermediate [%]
END_VAR
VAR CONSTANT
    DL_TR_MAX_RATE : REAL := 1000.0;           // 变化率上限 [%/s] / rate upper bound [%/s]
    DL_TR_MIN_RATE : REAL := 0.01;             // 变化率下限 [%/s] / rate lower bound [%/s]
    DL_TR_OUT_LIM  : REAL := 100.0;            // 输出双侧限幅 [%] / symmetrical output limit [%]
    DL_TR_DT       : TIME := T#10MS;           // 假定的任务周期，必须与实际一致 [ms] / assumed task period, must match the real one [ms]
    DL_TR_MS_SEC   : REAL := 1000.0;           // 毫秒转秒的除数，恒非零 [ms/s] / milliseconds to seconds divisor, never zero [ms/s]
    DL_FLOAT_EPS   : REAL := 1.0E-6;           // 浮点判等容差 [%] / float equality tolerance [%]
    DL_TR_INF_GUARD: REAL := 4.0E38;           // 非有限幅值判定阈值 [%] / non-finite magnitude guard [%]
    DL_TR_ZERO     : REAL := 0.0;              // 零值常量，避免裸字面量 [无量纲] / zero constant, avoids a bare literal [dimensionless]
END_VAR

// 段 1｜边沿实例无条件周期刷新（红线：严禁放入条件分支）/ segment 1, unconditional edge refresh
fbTrigReset(CLK := bReset);

// 段 2｜输出与错误状态预置 / segment 2, preset outputs and error status
eErr := 0;                                     // 预置无错误 / preset no error
bError := FALSE;                               // 预置无故障 / preset no fault
bTracking := FALSE;                            // 默认非跟踪态 / default not tracking
bInTransfer := FALSE;                          // 默认非过渡态 / default not transferring
tDelta := DL_TR_DT;                            // 本拍时间增量取固定任务周期 / this cycle increment uses the fixed task period

// 段 3｜首扫初始化（初值 FALSE，判据 NOT bInit）/ segment 3, first-scan initialisation
IF NOT bInit THEN
    eState := E_DL_TransferState.eIdle;        // 首扫落空闲态 / start in the idle state
    fLastOut := DL_TR_ZERO;                    // 输出记忆清零 / clear the output memory
    tLast := T#0MS;                            // 过渡时长清零 / clear the transfer time
    bInit := TRUE;                             // 首扫只做一次 / first scan runs once only
END_IF

// 段 4｜使能闸：失能输出 0 并清过渡 / segment 4, enable gate zeroes the output
IF NOT bEnable THEN
    eState := E_DL_TransferState.eIdle;        // 回空闲态 / back to idle
    fLastOut := DL_TR_ZERO;                    // 清输出记忆 / clear the output memory
    tLast := T#0MS;                            // 清过渡时长 / clear the transfer time
    fOut := DL_TR_ZERO;                        // 输出 0 / output zero
    fDeviation := DL_TR_ZERO;                  // 偏差 0 / deviation zero
    tInTransfer := T#0MS;                      // 过渡时长 0 / transfer time zero
    RETURN;                                    // 失能即出口 / disabled is the exit
END_IF

// 段 5｜斜率参数闸：非法即禁用过渡并直接取 PID 输出 / segment 5, rate parameter gate
bRateOk := (fRateMax >= DL_TR_MIN_RATE) AND (fRateMax <= DL_TR_MAX_RATE); // 域判定用与逻辑 / domain check by conjunction
IF NOT bRateOk THEN
    eErr := 16#0002_2410;                      // 斜率非法故障码 / illegal rate fault id
    bError := TRUE;                            // 置故障标志 / raise the error flag
END_IF

// 段 6｜给定非有限闸：任一给定非有限即落故障态，保持末次输出 / segment 6, non-finite setpoint gate
bNonFin := (fPidOut <> fPidOut) OR (fPidOut > DL_TR_INF_GUARD) OR (fPidOut < -DL_TR_INF_GUARD)
        OR (fTrackVal <> fTrackVal) OR (fTrackVal > DL_TR_INF_GUARD) OR (fTrackVal < -DL_TR_INF_GUARD)
        OR (fManualOut <> fManualOut) OR (fManualOut > DL_TR_INF_GUARD) OR (fManualOut < -DL_TR_INF_GUARD); // 三路给定同口径检查 / all three setpoints checked the same way
IF bNonFin THEN
    eErr := 16#0002_2411;                      // 给定非有限故障码 / non-finite setpoint fault id
    bError := TRUE;                            // 置故障标志 / raise the error flag
    eState := E_DL_TransferState.eFault;       // 落故障态 / enter the fault state
END_IF

// 段 7｜复位沿处理：放弃过渡，直接取目标值 / segment 7, reset abandons the transfer
IF fbTrigReset.Q THEN
    tLast := T#0MS;                            // 清过渡时长 / clear the transfer time
    IF bAuto THEN
        eState := E_DL_TransferState.eAuto;    // 直接进自动态 / jump straight to auto
        fLastOut := fPidOut;                   // 直接取 PID 输出 / take the PID output directly
    ELSE
        eState := E_DL_TransferState.eManual;  // 回手动态 / back to manual
        fLastOut := fTrackVal;                 // 取跟踪目标 / take the tracking target
    END_IF
END_IF

// 段 8｜单拍步长：斜率乘秒数，斜率已过闸，除数为常量恒非零 / segment 8, per cycle step size
IF bRateOk THEN
    fStep := fRateMax * TIME_TO_REAL(tDelta) / DL_TR_MS_SEC; // 步长 [%] / step size in percent
ELSE
    fStep := DL_TR_ZERO;                       // 斜率非法时步长 0，过渡不启用 / invalid rate yields a zero step, the transfer stays disabled
END_IF

// 段 9｜状态机主体（CASE 必含 ELSE 兜底，红线）/ segment 9, state machine body
CASE eState OF
    E_DL_TransferState.eIdle :
        fLastOut := DL_TR_ZERO;                // 空闲态输出记忆为 0 / the idle state keeps a zero output memory
        tLast := T#0MS;                        // 过渡时长清零 / clear the transfer time
        IF bAuto THEN
            eState := E_DL_TransferState.eTransfer; // 已请求自动，直接进过渡 / auto requested, enter the transfer
        ELSE
            eState := E_DL_TransferState.eManual;   // 否则进手动跟踪 / otherwise enter manual tracking
        END_IF
    E_DL_TransferState.eManual :
        bTracking := TRUE;                     // 手动期跟踪标志 / tracking flag in manual mode
        fClamped := MIN(MAX(fTrackVal, -DL_TR_OUT_LIM), DL_TR_OUT_LIM); // 手动期输出跟踪实际反馈，双侧限幅 / manual output tracks the actual feedback, clamped both sides
        fLastOut := fClamped;                  // 更新输出记忆 / update the output memory
        tLast := T#0MS;                        // 过渡时长清零，接管时从 0 计时 / clear the transfer time, counted from zero on takeover
        IF bAuto THEN
            eState := E_DL_TransferState.eTransfer; // 自动请求到来即进入过渡 / an auto request starts the transfer
        END_IF
    E_DL_TransferState.eTransfer :
        bInTransfer := TRUE;                   // 过渡进行中 / transfer in progress
        IF NOT bRateOk THEN
            fLastOut := fPidOut;               // 过渡禁用，直接取 PID 输出 / transfer disabled, take the PID output
            eState := E_DL_TransferState.eAuto;// 转自动态 / switch to auto
        ELSE
            tLast := tLast + tDelta;           // 累计过渡时长 / accumulate the transfer time
            IF ABS(fPidOut - fLastOut) <= (fStep + DL_FLOAT_EPS) THEN
                fLastOut := fPidOut;           // 收敛完成，落到 PID 输出 / converged, land on the PID output
                eState := E_DL_TransferState.eAuto; // 转自动态 / switch to auto
            ELSIF fPidOut > fLastOut THEN
                fLastOut := fLastOut + fStep;  // 正向逼近一个步长 / approach upwards by one step
            ELSE
                fLastOut := fLastOut - fStep;  // 负向逼近一个步长 / approach downwards by one step
            END_IF
            IF ABS(fPidOut - fLastOut) > fDevWindow THEN
                eErr := 16#0002_2401;          // 偏差超提示窗（信息级不置故障）/ deviation above the hint window, info level never raises a fault
            END_IF
        END_IF
        IF NOT bAuto THEN
            eState := E_DL_TransferState.eManual; // 中途撤回自动，回手动跟踪 / auto revoked mid-flight, back to manual tracking
            tLast := T#0MS;                    // 过渡时长清零 / clear the transfer time
        END_IF
    E_DL_TransferState.eAuto :
        fLastOut := fPidOut;                   // 自动态输出等于 PID 输出 / in auto the output equals the PID output
        tLast := T#0MS;                        // 过渡结束，时长清零 / transfer finished, clear the time
        IF NOT bAuto THEN
            eState := E_DL_TransferState.eManual; // 手动请求，回跟踪态 / a manual request returns to tracking
        END_IF
    E_DL_TransferState.eFault :
        bInTransfer := FALSE;                  // 故障态不过渡 / no transfer in the fault state
        fLastOut := MIN(MAX(fLastOut, -DL_TR_OUT_LIM), DL_TR_OUT_LIM); // 故障态保持末次输出，仅双侧限幅 / the fault state holds the last output, clamped both sides only
ELSE
    eErr := 16#0002_2411;                      // 非法状态兜底码，与给定非有限共用同一业务语义 / fallback code sharing the business meaning of a non-finite setpoint
    bError := TRUE;                            // 置故障标志 / raise the error flag
    eState := E_DL_TransferState.eFault;       // 一律回安全故障态 / always fall back to the safe fault state
    bInTransfer := FALSE;                      // 清除过渡标志 / clear the transfer flag
END_CASE

// 段 10｜输出双侧限幅与偏差监视 / segment 10, symmetrical clamping and deviation monitoring
fClamped := MIN(MAX(fLastOut, -DL_TR_OUT_LIM), DL_TR_OUT_LIM); // 双侧限幅，绝不只做单侧 / clamp both sides, never one side only
fOut := fClamped;                              // 输出镜像 / publish the output
fDeviation := fPidOut - fClamped;              // 偏差按限幅后的实际输出计算 / the deviation uses the clamped actual output
tInTransfer := tLast;                          // 过渡时长镜像 / publish the transfer time
END_FUNCTION_BLOCK
